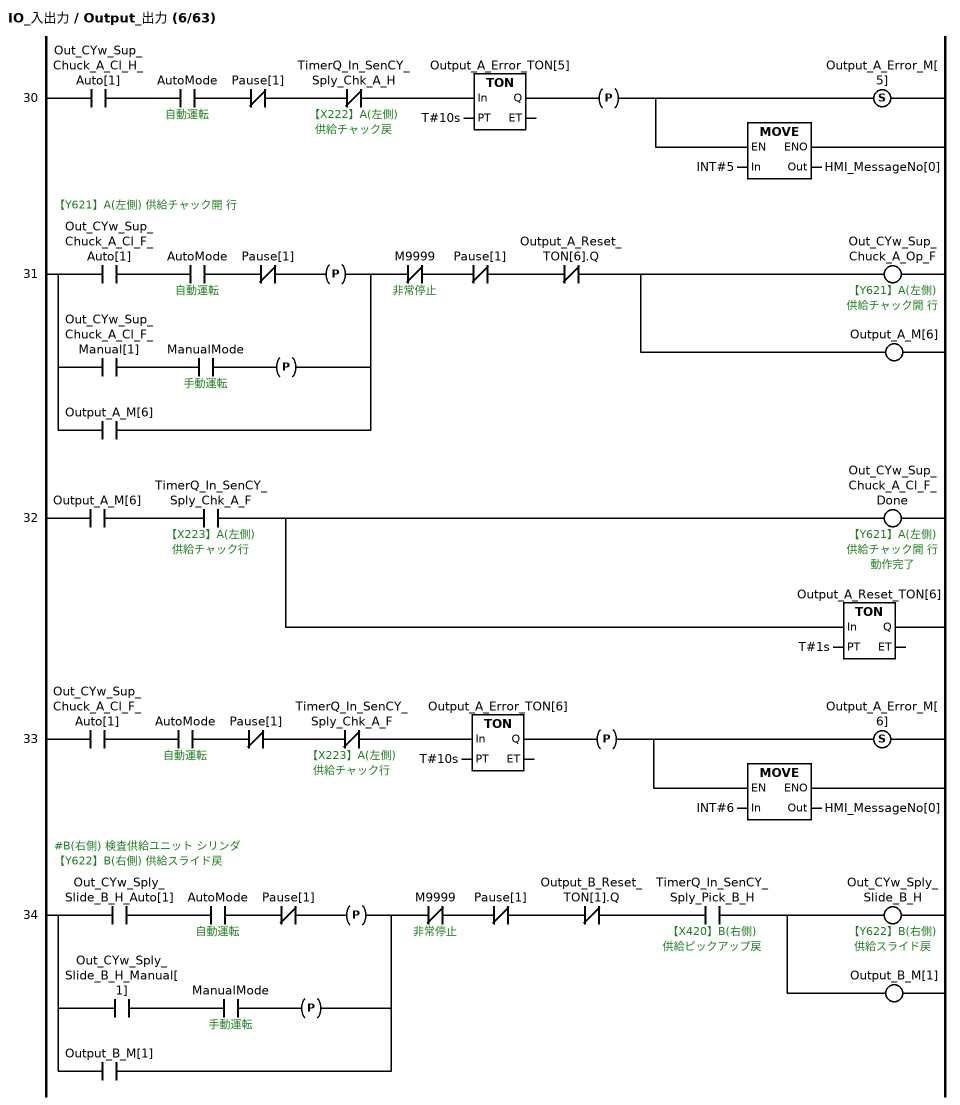
(* [picture p74: IO_入出力 / Output_出力, rungs 30-34] *)
(* Rung 30 *)
Output_A_Error_TON[5](In := Out_CYw_Sup_Chuck_A_Cl_H_Auto[1] AND AutoMode AND NOT Pause[1] AND NOT TimerQ_In_SenCY_Sply_Chk_A_H, PT := T#10s);
_e20(CLK := Output_A_Error_TON[5].Q);
IF _e20.Q THEN
    Output_A_Error_M[5] := TRUE;
    HMI_MessageNo[0] := INT#5;
END_IF;
(* Rung 31: 【Y621】A(左側) 供給チャック開 行 *)
_e21(CLK := Out_CYw_Sup_Chuck_A_Cl_F_Auto[1] AND AutoMode AND NOT Pause[1]);
_e22(CLK := Out_CYw_Sup_Chuck_A_Cl_F_Manual[1] AND ManualMode);
_p23 := (_e21.Q OR _e22.Q OR Output_A_M[6]) AND NOT M9999 AND NOT Pause[1] AND NOT Output_A_Reset_TON[6].Q;
Out_CYw_Sup_Chuck_A_Op_F := _p23;
Output_A_M[6] := _p23;
(* Rung 32 *)
Out_CYw_Sup_Chuck_A_Cl_F_Done := Output_A_M[6] AND TimerQ_In_SenCY_Sply_Chk_A_F;
Output_A_Reset_TON[6](In := Output_A_M[6] AND TimerQ_In_SenCY_Sply_Chk_A_F, PT := T#1s);
(* Rung 33 *)
Output_A_Error_TON[6](In := Out_CYw_Sup_Chuck_A_Cl_F_Auto[1] AND AutoMode AND NOT Pause[1] AND NOT TimerQ_In_SenCY_Sply_Chk_A_F, PT := T#10s);
_e24(CLK := Output_A_Error_TON[6].Q);
IF _e24.Q THEN
    Output_A_Error_M[6] := TRUE;
    HMI_MessageNo[0] := INT#6;
END_IF;
(* Rung 34: #B(右側) 検査供給ユニット シリンダ / 【Y622】B(右側) 供給スライド戻 *)
_e25(CLK := Out_CYw_Sply_Slide_B_H_Auto[1] AND AutoMode AND NOT Pause[1]);
_e26(CLK := Out_CYw_Sply_Slide_B_H_Manual[1] AND ManualMode);
_p27 := (_e25.Q OR _e26.Q OR Output_B_M[1]) AND NOT M9999 AND NOT Pause[1] AND NOT Output_B_Reset_TON[1].Q AND TimerQ_In_SenCY_Sply_Pick_B_H;
Out_CYw_Sply_Slide_B_H := _p27;
Output_B_M[1] := _p27;

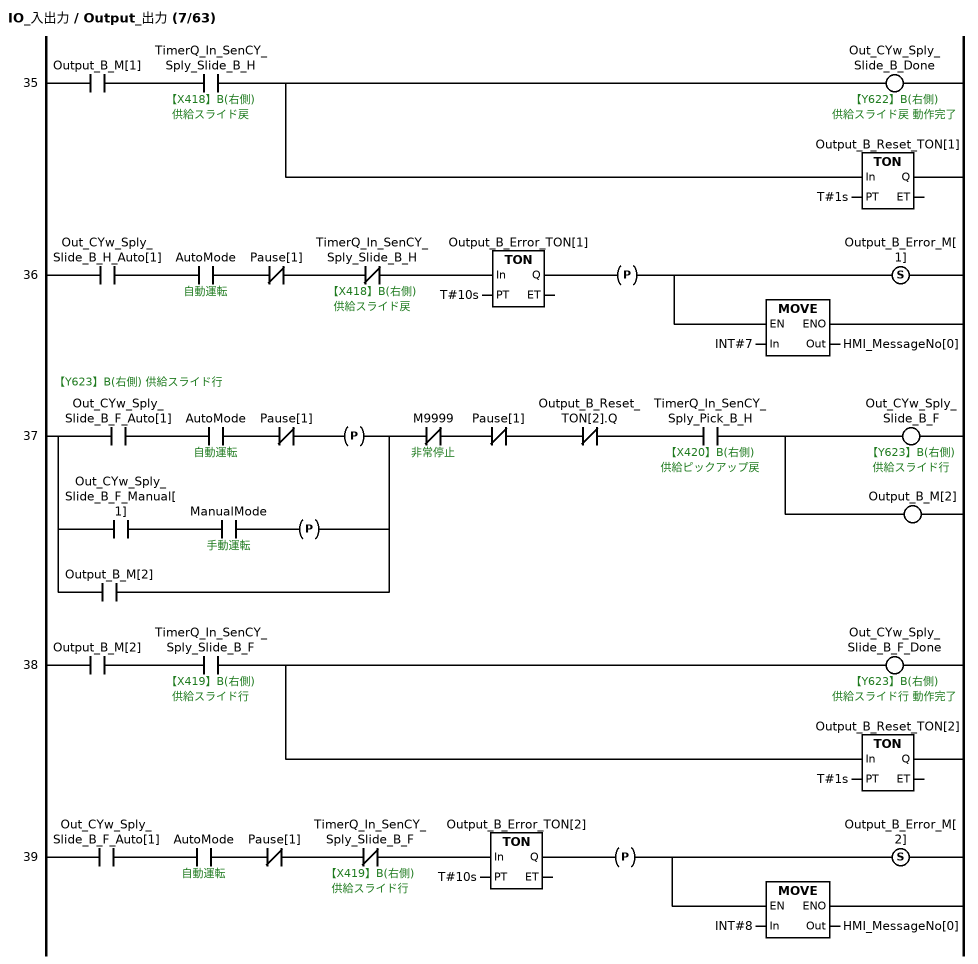
(* Rung 35 *)
Out_CYw_Sply_Slide_B_Done := Output_B_M[1] AND TimerQ_In_SenCY_Sply_Slide_B_H;
Output_B_Reset_TON[1](In := Output_B_M[1] AND TimerQ_In_SenCY_Sply_Slide_B_H, PT := T#1s);
(* Rung 36 *)
Output_B_Error_TON[1](In := Out_CYw_Sply_Slide_B_H_Auto[1] AND AutoMode AND NOT Pause[1] AND NOT TimerQ_In_SenCY_Sply_Slide_B_H, PT := T#10s);
_e28(CLK := Output_B_Error_TON[1].Q);
IF _e28.Q THEN
    Output_B_Error_M[1] := TRUE;
    HMI_MessageNo[0] := INT#7;
END_IF;
(* Rung 37: 【Y623】B(右側) 供給スライド行 *)
_e29(CLK := Out_CYw_Sply_Slide_B_F_Auto[1] AND AutoMode AND NOT Pause[1]);
_e30(CLK := Out_CYw_Sply_Slide_B_F_Manual[1] AND ManualMode);
_p31 := (_e29.Q OR _e30.Q OR Output_B_M[2]) AND NOT M9999 AND NOT Pause[1] AND NOT Output_B_Reset_TON[2].Q AND TimerQ_In_SenCY_Sply_Pick_B_H;
Out_CYw_Sply_Slide_B_F := _p31;
Output_B_M[2] := _p31;
(* Rung 38 *)
Out_CYw_Sply_Slide_B_F_Done := Output_B_M[2] AND TimerQ_In_SenCY_Sply_Slide_B_F;
Output_B_Reset_TON[2](In := Output_B_M[2] AND TimerQ_In_SenCY_Sply_Slide_B_F, PT := T#1s);
(* Rung 39 *)
Output_B_Error_TON[2](In := Out_CYw_Sply_Slide_B_F_Auto[1] AND AutoMode AND NOT Pause[1] AND NOT TimerQ_In_SenCY_Sply_Slide_B_F, PT := T#10s);
_e32(CLK := Output_B_Error_TON[2].Q);
IF _e32.Q THEN
    Output_B_Error_M[2] := TRUE;
    HMI_MessageNo[0] := INT#8;
END_IF;

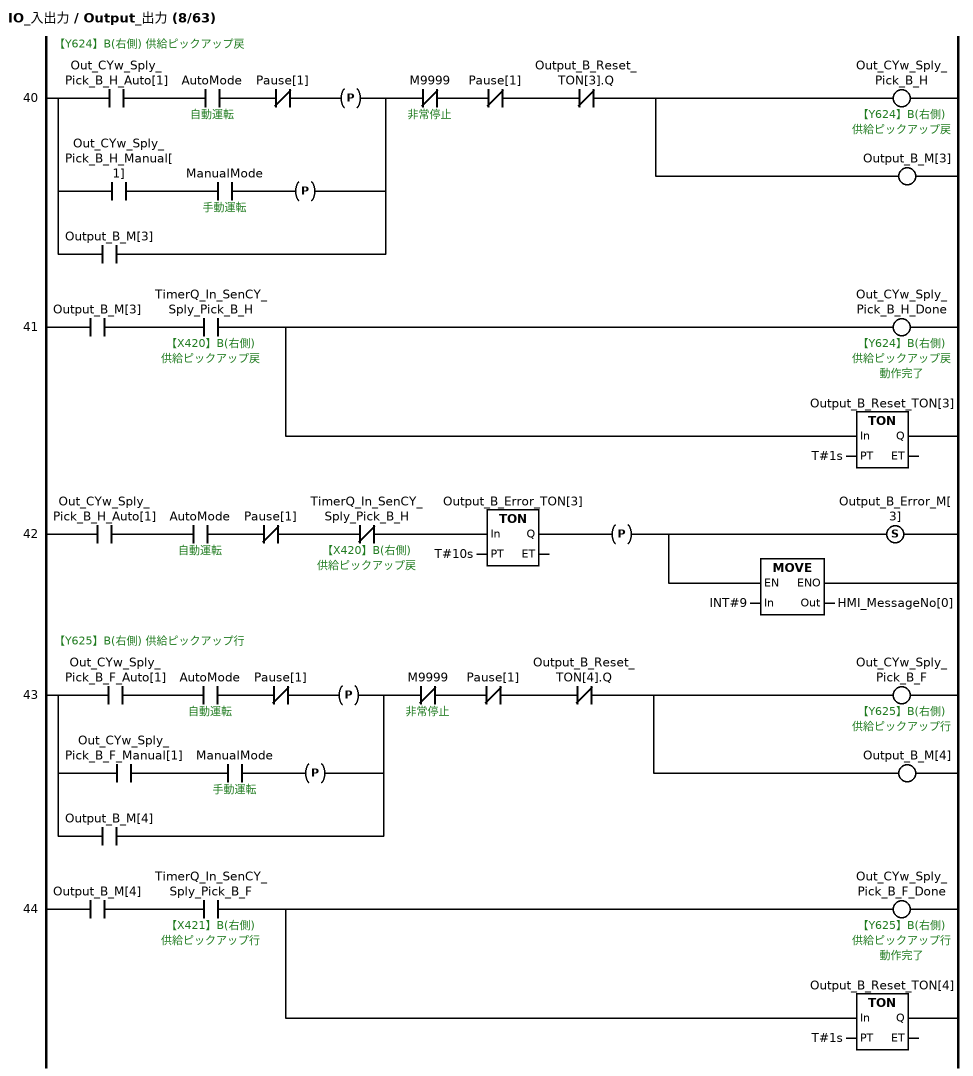
(* Rung 40: 【Y624】B(右側) 供給ピックアップ戻 *)
_e33(CLK := Out_CYw_Sply_Pick_B_H_Auto[1] AND AutoMode AND NOT Pause[1]);
_e34(CLK := Out_CYw_Sply_Pick_B_H_Manual[1] AND ManualMode);
_p35 := (_e33.Q OR _e34.Q OR Output_B_M[3]) AND NOT M9999 AND NOT Pause[1] AND NOT Output_B_Reset_TON[3].Q;
Out_CYw_Sply_Pick_B_H := _p35;
Output_B_M[3] := _p35;
(* Rung 41 *)
Out_CYw_Sply_Pick_B_H_Done := Output_B_M[3] AND TimerQ_In_SenCY_Sply_Pick_B_H;
Output_B_Reset_TON[3](In := Output_B_M[3] AND TimerQ_In_SenCY_Sply_Pick_B_H, PT := T#1s);
(* Rung 42 *)
Output_B_Error_TON[3](In := Out_CYw_Sply_Pick_B_H_Auto[1] AND AutoMode AND NOT Pause[1] AND NOT TimerQ_In_SenCY_Sply_Pick_B_H, PT := T#10s);
_e36(CLK := Output_B_Error_TON[3].Q);
IF _e36.Q THEN
    Output_B_Error_M[3] := TRUE;
    HMI_MessageNo[0] := INT#9;
END_IF;
(* Rung 43: 【Y625】B(右側) 供給ピックアップ行 *)
_e37(CLK := Out_CYw_Sply_Pick_B_F_Auto[1] AND AutoMode AND NOT Pause[1]);
_e38(CLK := Out_CYw_Sply_Pick_B_F_Manual[1] AND ManualMode);
_p39 := (_e37.Q OR _e38.Q OR Output_B_M[4]) AND NOT M9999 AND NOT Pause[1] AND NOT Output_B_Reset_TON[4].Q;
Out_CYw_Sply_Pick_B_F := _p39;
Output_B_M[4] := _p39;
(* Rung 44 *)
Out_CYw_Sply_Pick_B_F_Done := Output_B_M[4] AND TimerQ_In_SenCY_Sply_Pick_B_F;
Output_B_Reset_TON[4](In := Output_B_M[4] AND TimerQ_In_SenCY_Sply_Pick_B_F, PT := T#1s);

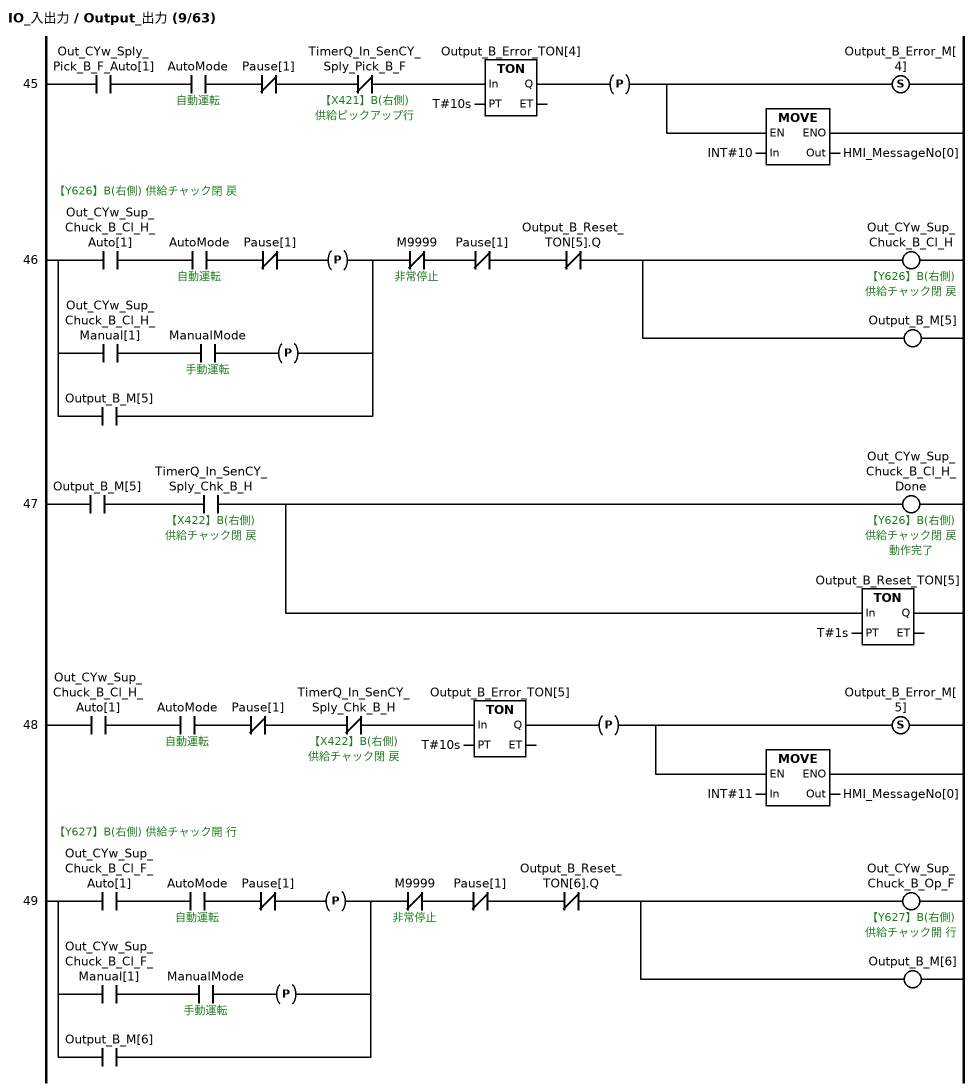
(* Rung 45 *)
Output_B_Error_TON[4](In := Out_CYw_Sply_Pick_B_F_Auto[1] AND AutoMode AND NOT Pause[1] AND NOT TimerQ_In_SenCY_Sply_Pick_B_F, PT := T#10s);
_e40(CLK := Output_B_Error_TON[4].Q);
IF _e40.Q THEN
    Output_B_Error_M[4] := TRUE;
    HMI_MessageNo[0] := INT#10;
END_IF;
(* Rung 46: 【Y626】B(右側) 供給チャック閉 戻 *)
_e41(CLK := Out_CYw_Sup_Chuck_B_Cl_H_Auto[1] AND AutoMode AND NOT Pause[1]);
_e42(CLK := Out_CYw_Sup_Chuck_B_Cl_H_Manual[1] AND ManualMode);
_p43 := (_e41.Q OR _e42.Q OR Output_B_M[5]) AND NOT M9999 AND NOT Pause[1] AND NOT Output_B_Reset_TON[5].Q;
Out_CYw_Sup_Chuck_B_Cl_H := _p43;
Output_B_M[5] := _p43;
(* Rung 47 *)
Out_CYw_Sup_Chuck_B_Cl_H_Done := Output_B_M[5] AND TimerQ_In_SenCY_Sply_Chk_B_H;
Output_B_Reset_TON[5](In := Output_B_M[5] AND TimerQ_In_SenCY_Sply_Chk_B_H, PT := T#1s);
(* Rung 48 *)
Output_B_Error_TON[5](In := Out_CYw_Sup_Chuck_B_Cl_H_Auto[1] AND AutoMode AND NOT Pause[1] AND NOT TimerQ_In_SenCY_Sply_Chk_B_H, PT := T#10s);
_e44(CLK := Output_B_Error_TON[5].Q);
IF _e44.Q THEN
    Output_B_Error_M[5] := TRUE;
    HMI_MessageNo[0] := INT#11;
END_IF;
(* Rung 49: 【Y627】B(右側) 供給チャック開 行 *)
_e45(CLK := Out_CYw_Sup_Chuck_B_Cl_F_Auto[1] AND AutoMode AND NOT Pause[1]);
_e46(CLK := Out_CYw_Sup_Chuck_B_Cl_F_Manual[1] AND ManualMode);
_p47 := (_e45.Q OR _e46.Q OR Output_B_M[6]) AND NOT M9999 AND NOT Pause[1] AND NOT Output_B_Reset_TON[6].Q;
Out_CYw_Sup_Chuck_B_Op_F := _p47;
Output_B_M[6] := _p47;

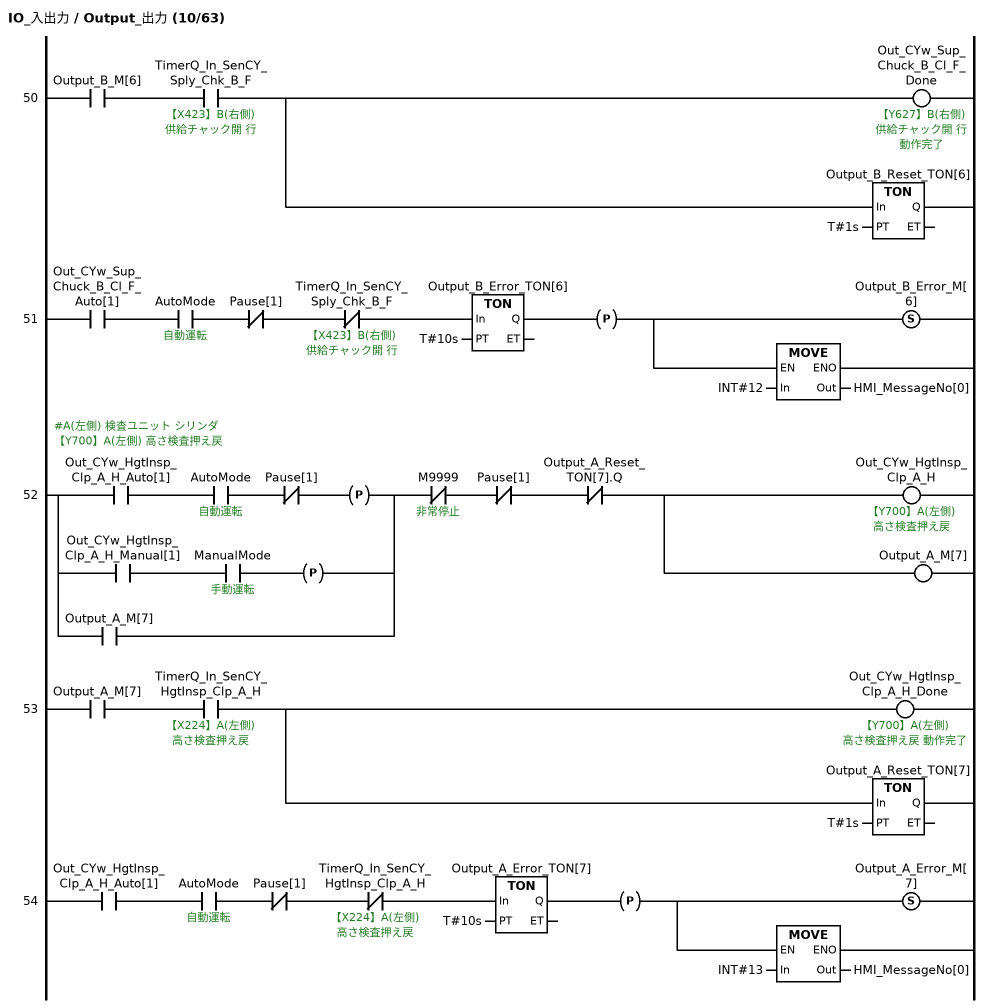
(* Rung 50 *)
Out_CYw_Sup_Chuck_B_Cl_F_Done := Output_B_M[6] AND TimerQ_In_SenCY_Sply_Chk_B_F;
Output_B_Reset_TON[6](In := Output_B_M[6] AND TimerQ_In_SenCY_Sply_Chk_B_F, PT := T#1s);
(* Rung 51 *)
Output_B_Error_TON[6](In := Out_CYw_Sup_Chuck_B_Cl_F_Auto[1] AND AutoMode AND NOT Pause[1] AND NOT TimerQ_In_SenCY_Sply_Chk_B_F, PT := T#10s);
_e48(CLK := Output_B_Error_TON[6].Q);
IF _e48.Q THEN
    Output_B_Error_M[6] := TRUE;
    HMI_MessageNo[0] := INT#12;
END_IF;
(* Rung 52: #A(左側) 検査ユニット シリンダ / 【Y700】A(左側) 高さ検査押え戻 *)
_e49(CLK := Out_CYw_HgtInsp_Clp_A_H_Auto[1] AND AutoMode AND NOT Pause[1]);
_e50(CLK := Out_CYw_HgtInsp_Clp_A_H_Manual[1] AND ManualMode);
_p51 := (_e49.Q OR _e50.Q OR Output_A_M[7]) AND NOT M9999 AND NOT Pause[1] AND NOT Output_A_Reset_TON[7].Q;
Out_CYw_HgtInsp_Clp_A_H := _p51;
Output_A_M[7] := _p51;
(* Rung 53 *)
_p52 := Output_A_M[7] AND TimerQ_In_SenCY_HgtInsp_Clp_A_H;
Out_CYw_HgtInsp_Clp_A_H_Done := _p52;
Output_A_Reset_TON[7](In := _p52, PT := T#1s);
(* Rung 54 *)
Output_A_Error_TON[7](In := Out_CYw_HgtInsp_Clp_A_H_Auto[1] AND AutoMode AND NOT Pause[1] AND NOT TimerQ_In_SenCY_HgtInsp_Clp_A_H, PT := T#10s);
_e53(CLK := Output_A_Error_TON[7].Q);
IF _e53.Q THEN
    Output_A_Error_M[7] := TRUE;
    HMI_MessageNo[0] := INT#13;
END_IF;

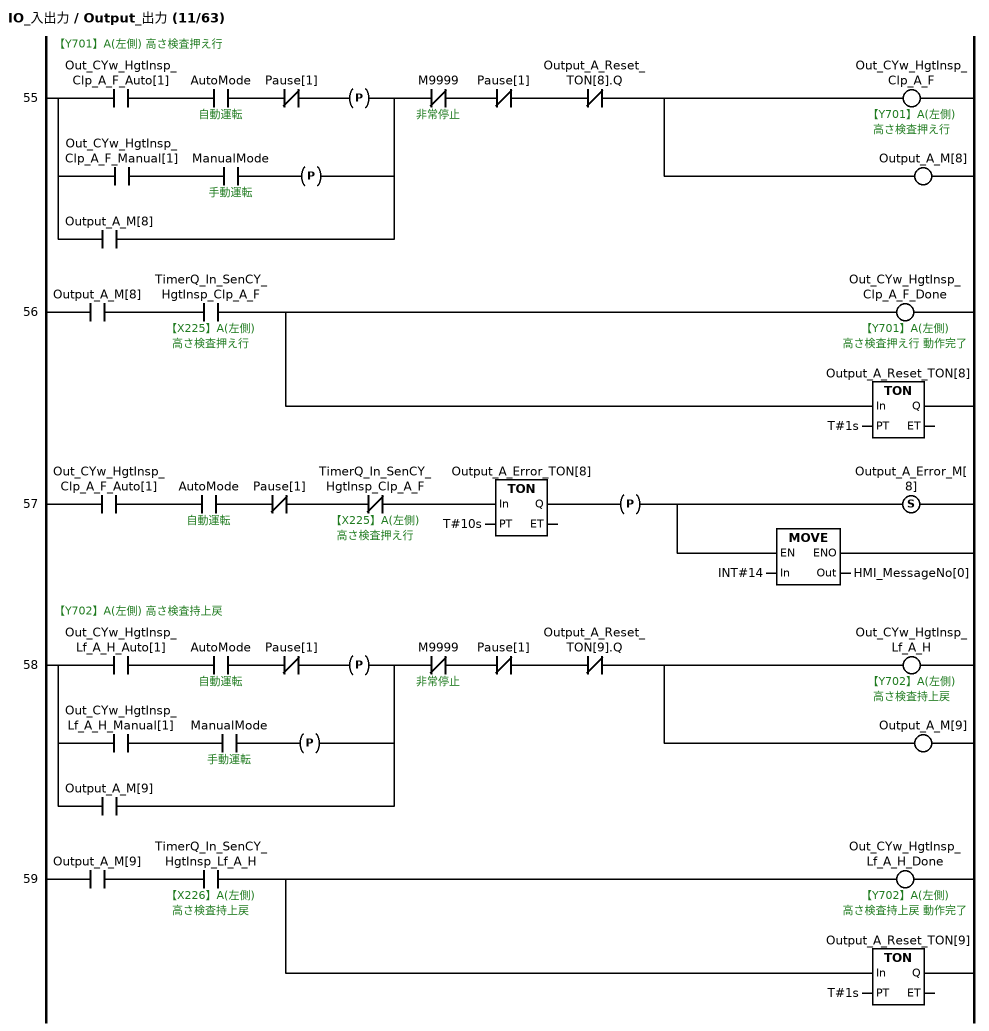
(* Rung 55: 【Y701】A(左側) 高さ検査押え行 *)
_e54(CLK := Out_CYw_HgtInsp_Clp_A_F_Auto[1] AND AutoMode AND NOT Pause[1]);
_e55(CLK := Out_CYw_HgtInsp_Clp_A_F_Manual[1] AND ManualMode);
_p56 := (_e54.Q OR _e55.Q OR Output_A_M[8]) AND NOT M9999 AND NOT Pause[1] AND NOT Output_A_Reset_TON[8].Q;
Out_CYw_HgtInsp_Clp_A_F := _p56;
Output_A_M[8] := _p56;
(* Rung 56 *)
_p57 := Output_A_M[8] AND TimerQ_In_SenCY_HgtInsp_Clp_A_F;
Out_CYw_HgtInsp_Clp_A_F_Done := _p57;
Output_A_Reset_TON[8](In := _p57, PT := T#1s);
(* Rung 57 *)
Output_A_Error_TON[8](In := Out_CYw_HgtInsp_Clp_A_F_Auto[1] AND AutoMode AND NOT Pause[1] AND NOT TimerQ_In_SenCY_HgtInsp_Clp_A_F, PT := T#10s);
_e58(CLK := Output_A_Error_TON[8].Q);
IF _e58.Q THEN
    Output_A_Error_M[8] := TRUE;
    HMI_MessageNo[0] := INT#14;
END_IF;
(* Rung 58: 【Y702】A(左側) 高さ検査持上戻 *)
_e59(CLK := Out_CYw_HgtInsp_Lf_A_H_Auto[1] AND AutoMode AND NOT Pause[1]);
_e60(CLK := Out_CYw_HgtInsp_Lf_A_H_Manual[1] AND ManualMode);
_p61 := (_e59.Q OR _e60.Q OR Output_A_M[9]) AND NOT M9999 AND NOT Pause[1] AND NOT Output_A_Reset_TON[9].Q;
Out_CYw_HgtInsp_Lf_A_H := _p61;
Output_A_M[9] := _p61;
(* Rung 59 *)
Out_CYw_HgtInsp_Lf_A_H_Done := Output_A_M[9] AND TimerQ_In_SenCY_HgtInsp_Lf_A_H;
Output_A_Reset_TON[9](In := Output_A_M[9] AND TimerQ_In_SenCY_HgtInsp_Lf_A_H, PT := T#1s);

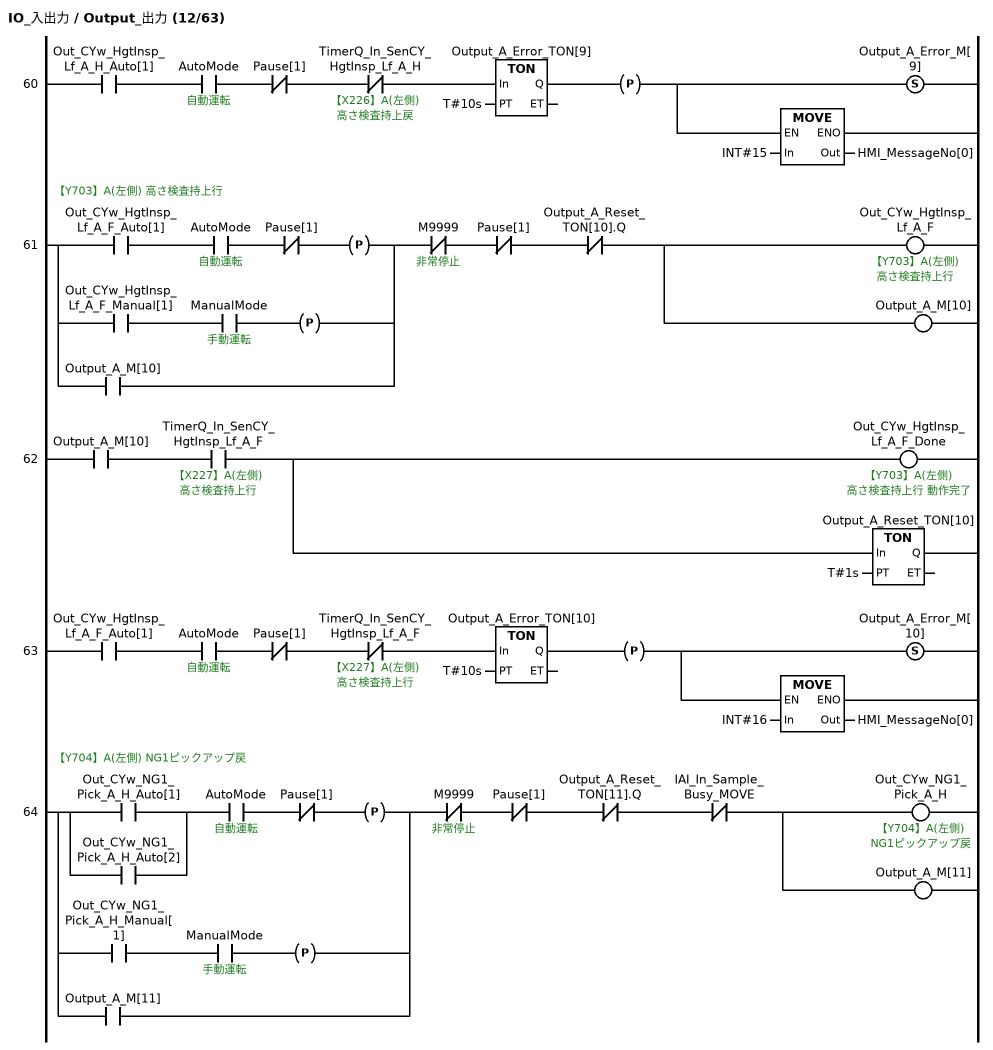
(* Rung 60 *)
Output_A_Error_TON[9](In := Out_CYw_HgtInsp_Lf_A_H_Auto[1] AND AutoMode AND NOT Pause[1] AND NOT TimerQ_In_SenCY_HgtInsp_Lf_A_H, PT := T#10s);
_e62(CLK := Output_A_Error_TON[9].Q);
IF _e62.Q THEN
    Output_A_Error_M[9] := TRUE;
    HMI_MessageNo[0] := INT#15;
END_IF;
(* Rung 61: 【Y703】A(左側) 高さ検査持上行 *)
_e63(CLK := Out_CYw_HgtInsp_Lf_A_F_Auto[1] AND AutoMode AND NOT Pause[1]);
_e64(CLK := Out_CYw_HgtInsp_Lf_A_F_Manual[1] AND ManualMode);
_p65 := (_e63.Q OR _e64.Q OR Output_A_M[10]) AND NOT M9999 AND NOT Pause[1] AND NOT Output_A_Reset_TON[10].Q;
Out_CYw_HgtInsp_Lf_A_F := _p65;
Output_A_M[10] := _p65;
(* Rung 62 *)
_p66 := Output_A_M[10] AND TimerQ_In_SenCY_HgtInsp_Lf_A_F;
Out_CYw_HgtInsp_Lf_A_F_Done := _p66;
Output_A_Reset_TON[10](In := _p66, PT := T#1s);
(* Rung 63 *)
Output_A_Error_TON[10](In := Out_CYw_HgtInsp_Lf_A_F_Auto[1] AND AutoMode AND NOT Pause[1] AND NOT TimerQ_In_SenCY_HgtInsp_Lf_A_F, PT := T#10s);
_e67(CLK := Output_A_Error_TON[10].Q);
IF _e67.Q THEN
    Output_A_Error_M[10] := TRUE;
    HMI_MessageNo[0] := INT#16;
END_IF;
(* Rung 64: 【Y704】A(左側) NG1ピックアップ戻 *)
_e68(CLK := (Out_CYw_NG1_Pick_A_H_Auto[1] OR Out_CYw_NG1_Pick_A_H_Auto[2]) AND AutoMode AND NOT Pause[1]);
_e69(CLK := Out_CYw_NG1_Pick_A_H_Manual[1] AND ManualMode);
_p70 := (_e68.Q OR _e69.Q OR Output_A_M[11]) AND NOT M9999 AND NOT Pause[1] AND NOT Output_A_Reset_TON[11].Q AND NOT IAI_In_Sample_Busy_MOVE;
Out_CYw_NG1_Pick_A_H := _p70;
Output_A_M[11] := _p70;

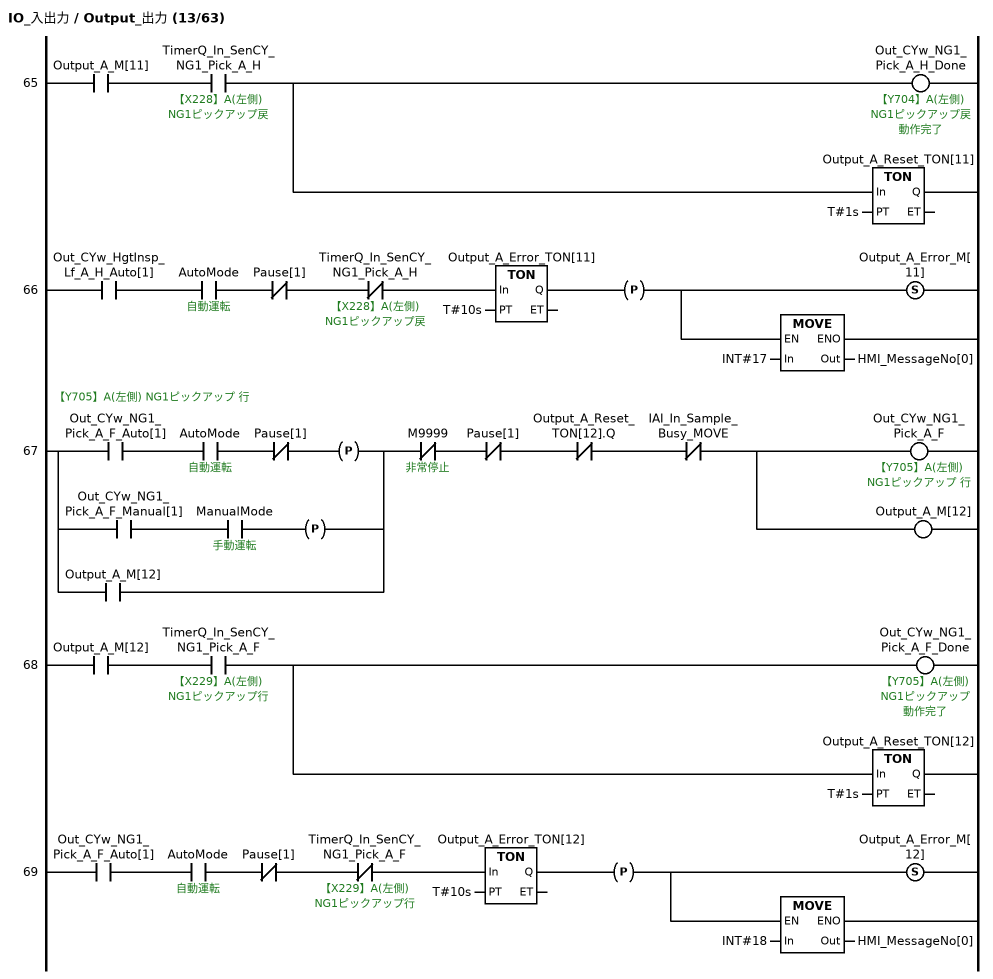
(* Rung 65 *)
Out_CYw_NG1_Pick_A_H_Done := Output_A_M[11] AND TimerQ_In_SenCY_NG1_Pick_A_H;
Output_A_Reset_TON[11](In := Output_A_M[11] AND TimerQ_In_SenCY_NG1_Pick_A_H, PT := T#1s);
(* Rung 66 *)
Output_A_Error_TON[11](In := Out_CYw_HgtInsp_Lf_A_H_Auto[1] AND AutoMode AND NOT Pause[1] AND NOT TimerQ_In_SenCY_NG1_Pick_A_H, PT := T#10s);
_e71(CLK := Output_A_Error_TON[11].Q);
IF _e71.Q THEN
    Output_A_Error_M[11] := TRUE;
    HMI_MessageNo[0] := INT#17;
END_IF;
(* Rung 67: 【Y705】A(左側) NG1ピックアップ 行 *)
_e72(CLK := Out_CYw_NG1_Pick_A_F_Auto[1] AND AutoMode AND NOT Pause[1]);
_e73(CLK := Out_CYw_NG1_Pick_A_F_Manual[1] AND ManualMode);
_p74 := (_e72.Q OR _e73.Q OR Output_A_M[12]) AND NOT M9999 AND NOT Pause[1] AND NOT Output_A_Reset_TON[12].Q AND NOT IAI_In_Sample_Busy_MOVE;
Out_CYw_NG1_Pick_A_F := _p74;
Output_A_M[12] := _p74;
(* Rung 68 *)
Out_CYw_NG1_Pick_A_F_Done := Output_A_M[12] AND TimerQ_In_SenCY_NG1_Pick_A_F;
Output_A_Reset_TON[12](In := Output_A_M[12] AND TimerQ_In_SenCY_NG1_Pick_A_F, PT := T#1s);
(* Rung 69 *)
Output_A_Error_TON[12](In := Out_CYw_NG1_Pick_A_F_Auto[1] AND AutoMode AND NOT Pause[1] AND NOT TimerQ_In_SenCY_NG1_Pick_A_F, PT := T#10s);
_e75(CLK := Output_A_Error_TON[12].Q);
IF _e75.Q THEN
    Output_A_Error_M[12] := TRUE;
    HMI_MessageNo[0] := INT#18;
END_IF;

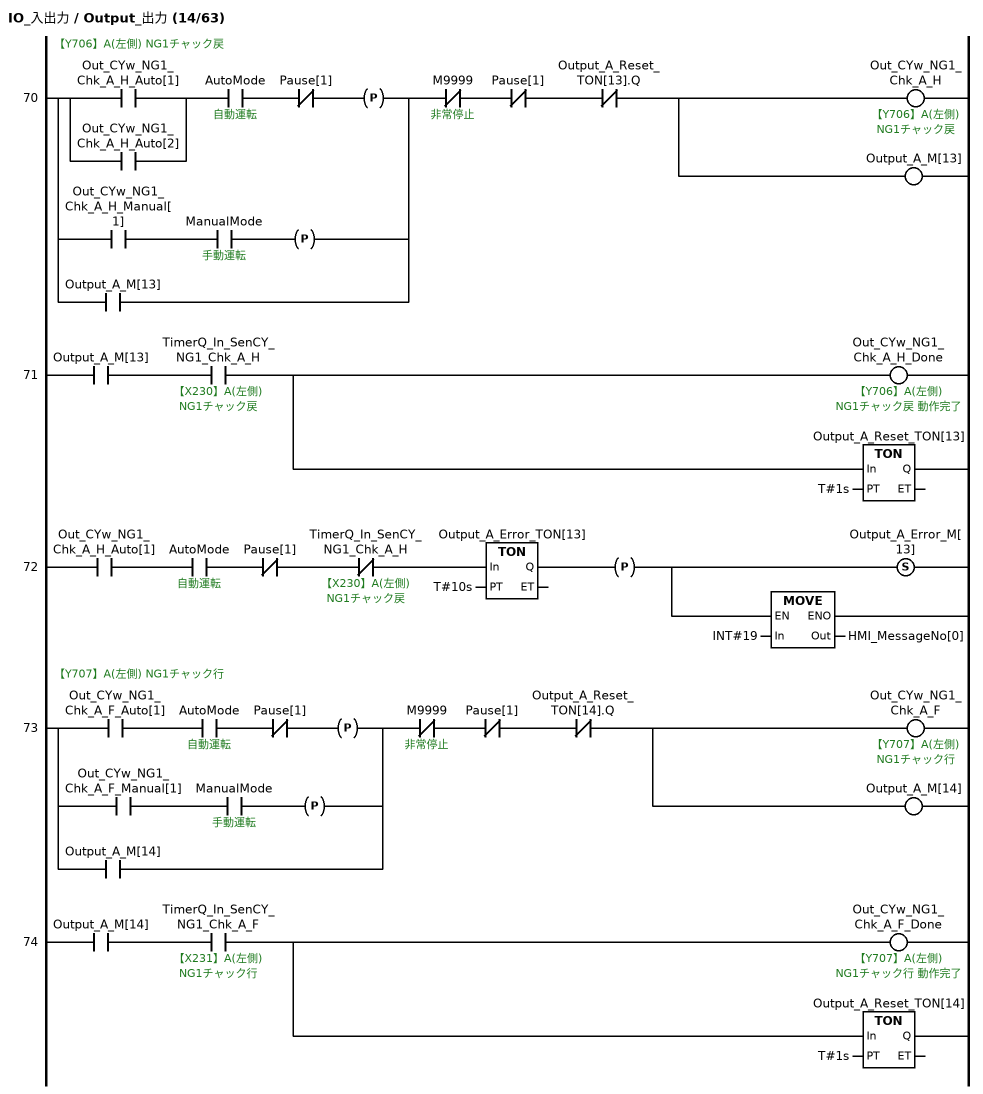
(* Rung 70: 【Y706】A(左側) NG1チャック戻 *)
_e76(CLK := (Out_CYw_NG1_Chk_A_H_Auto[1] OR Out_CYw_NG1_Chk_A_H_Auto[2]) AND AutoMode AND NOT Pause[1]);
_e77(CLK := Out_CYw_NG1_Chk_A_H_Manual[1] AND ManualMode);
_p78 := (_e76.Q OR _e77.Q OR Output_A_M[13]) AND NOT M9999 AND NOT Pause[1] AND NOT Output_A_Reset_TON[13].Q;
Out_CYw_NG1_Chk_A_H := _p78;
Output_A_M[13] := _p78;
(* Rung 71 *)
Out_CYw_NG1_Chk_A_H_Done := Output_A_M[13] AND TimerQ_In_SenCY_NG1_Chk_A_H;
Output_A_Reset_TON[13](In := Output_A_M[13] AND TimerQ_In_SenCY_NG1_Chk_A_H, PT := T#1s);
(* Rung 72 *)
Output_A_Error_TON[13](In := Out_CYw_NG1_Chk_A_H_Auto[1] AND AutoMode AND NOT Pause[1] AND NOT TimerQ_In_SenCY_NG1_Chk_A_H, PT := T#10s);
_e79(CLK := Output_A_Error_TON[13].Q);
IF _e79.Q THEN
    Output_A_Error_M[13] := TRUE;
    HMI_MessageNo[0] := INT#19;
END_IF;
(* Rung 73: 【Y707】A(左側) NG1チャック行 *)
_e80(CLK := Out_CYw_NG1_Chk_A_F_Auto[1] AND AutoMode AND NOT Pause[1]);
_e81(CLK := Out_CYw_NG1_Chk_A_F_Manual[1] AND ManualMode);
_p82 := (_e80.Q OR _e81.Q OR Output_A_M[14]) AND NOT M9999 AND NOT Pause[1] AND NOT Output_A_Reset_TON[14].Q;
Out_CYw_NG1_Chk_A_F := _p82;
Output_A_M[14] := _p82;
(* Rung 74 *)
Out_CYw_NG1_Chk_A_F_Done := Output_A_M[14] AND TimerQ_In_SenCY_NG1_Chk_A_F;
Output_A_Reset_TON[14](In := Output_A_M[14] AND TimerQ_In_SenCY_NG1_Chk_A_F, PT := T#1s);

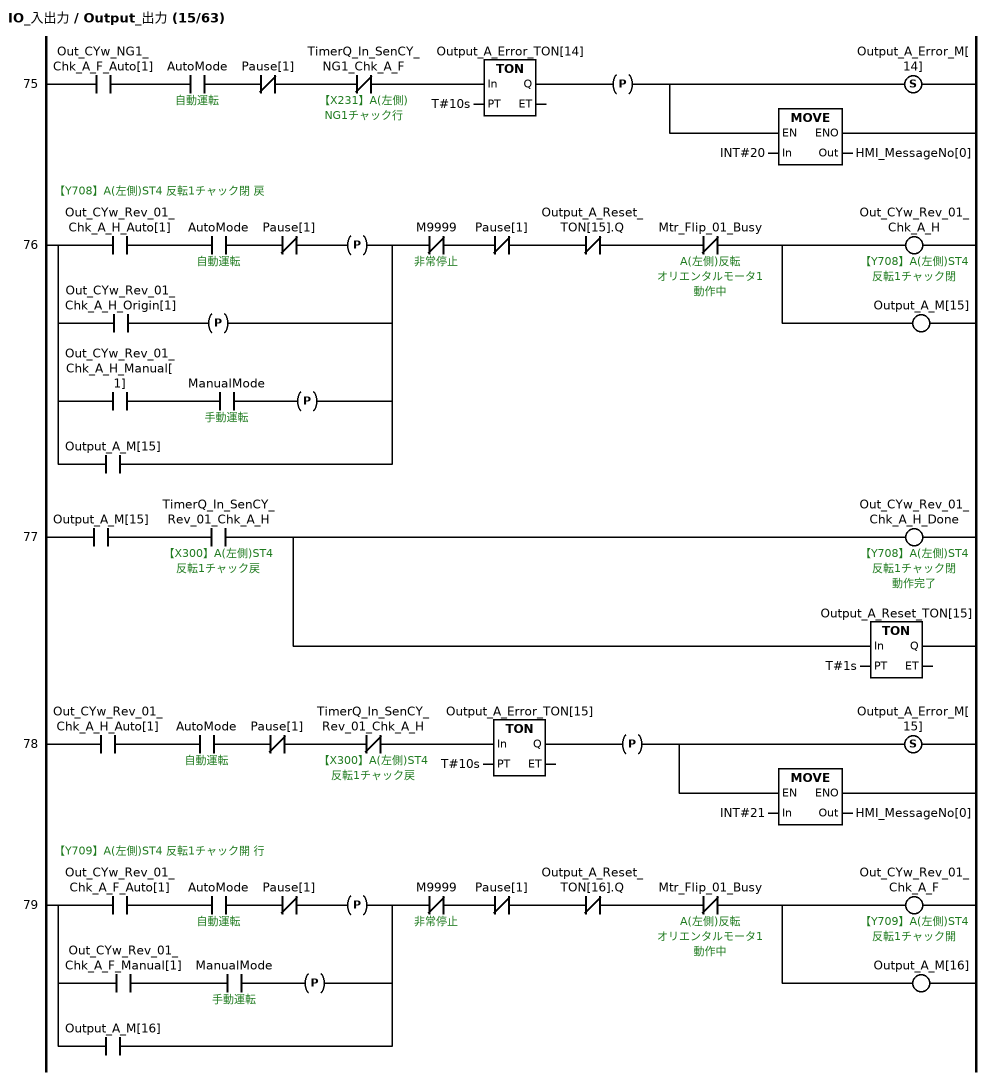
(* Rung 75 *)
Output_A_Error_TON[14](In := Out_CYw_NG1_Chk_A_F_Auto[1] AND AutoMode AND NOT Pause[1] AND NOT TimerQ_In_SenCY_NG1_Chk_A_F, PT := T#10s);
_e83(CLK := Output_A_Error_TON[14].Q);
IF _e83.Q THEN
    Output_A_Error_M[14] := TRUE;
    HMI_MessageNo[0] := INT#20;
END_IF;
(* Rung 76: 【Y708】A(左側)ST4 反転1チャック閉 戻 *)
_e84(CLK := Out_CYw_Rev_01_Chk_A_H_Auto[1] AND AutoMode AND NOT Pause[1]);
_e85(CLK := Out_CYw_Rev_01_Chk_A_H_Origin[1]);
_e86(CLK := Out_CYw_Rev_01_Chk_A_H_Manual[1] AND ManualMode);
_p87 := (_e84.Q OR _e85.Q OR _e86.Q OR Output_A_M[15]) AND NOT M9999 AND NOT Pause[1] AND NOT Output_A_Reset_TON[15].Q AND NOT Mtr_Flip_01_Busy;
Out_CYw_Rev_01_Chk_A_H := _p87;
Output_A_M[15] := _p87;
(* Rung 77 *)
_p88 := Output_A_M[15] AND TimerQ_In_SenCY_Rev_01_Chk_A_H;
Out_CYw_Rev_01_Chk_A_H_Done := _p88;
Output_A_Reset_TON[15](In := _p88, PT := T#1s);
(* Rung 78 *)
Output_A_Error_TON[15](In := Out_CYw_Rev_01_Chk_A_H_Auto[1] AND AutoMode AND NOT Pause[1] AND NOT TimerQ_In_SenCY_Rev_01_Chk_A_H, PT := T#10s);
_e89(CLK := Output_A_Error_TON[15].Q);
IF _e89.Q THEN
    Output_A_Error_M[15] := TRUE;
    HMI_MessageNo[0] := INT#21;
END_IF;
(* Rung 79: 【Y709】A(左側)ST4 反転1チャック開 行 *)
_e90(CLK := Out_CYw_Rev_01_Chk_A_F_Auto[1] AND AutoMode AND NOT Pause[1]);
_e91(CLK := Out_CYw_Rev_01_Chk_A_F_Manual[1] AND ManualMode);
_p92 := (_e90.Q OR _e91.Q OR Output_A_M[16]) AND NOT M9999 AND NOT Pause[1] AND NOT Output_A_Reset_TON[16].Q AND NOT Mtr_Flip_01_Busy;
Out_CYw_Rev_01_Chk_A_F := _p92;
Output_A_M[16] := _p92;

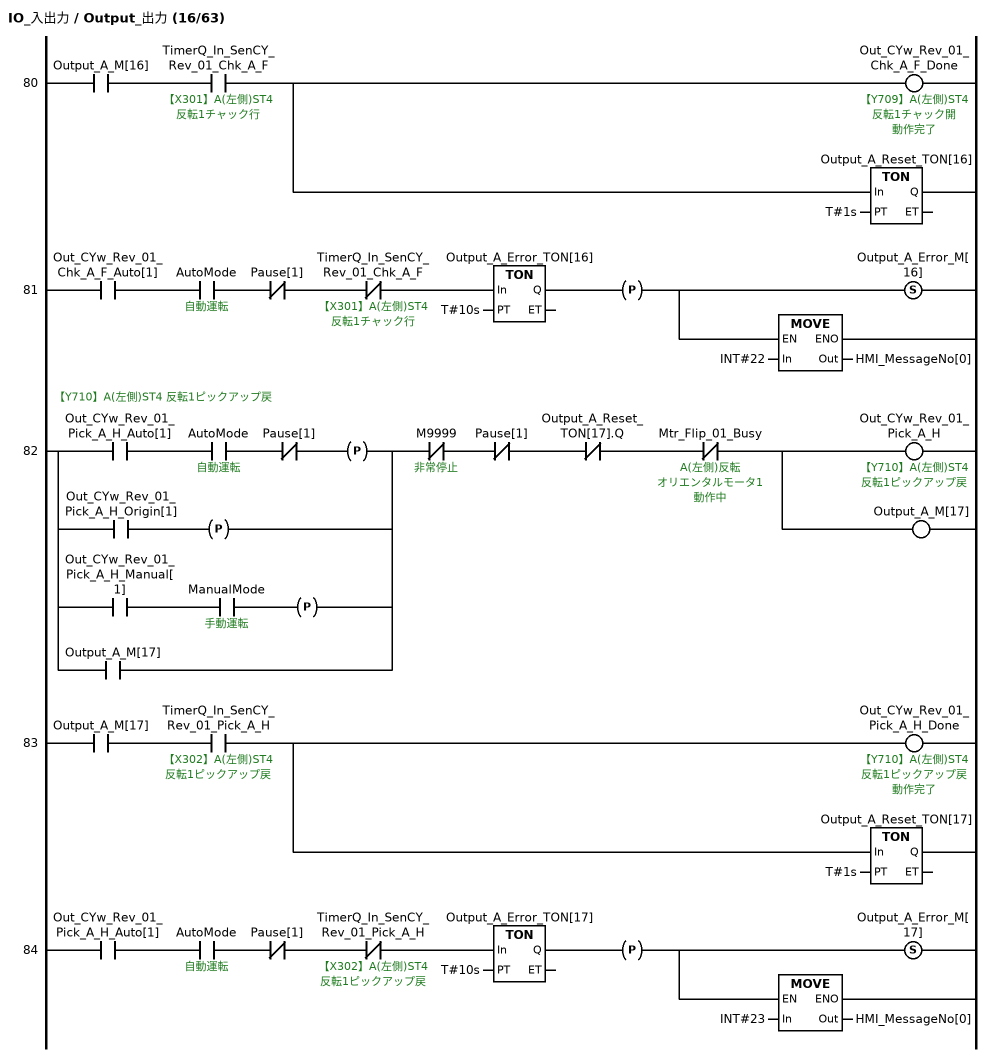
(* Rung 80 *)
_p93 := Output_A_M[16] AND TimerQ_In_SenCY_Rev_01_Chk_A_F;
Out_CYw_Rev_01_Chk_A_F_Done := _p93;
Output_A_Reset_TON[16](In := _p93, PT := T#1s);
(* Rung 81 *)
Output_A_Error_TON[16](In := Out_CYw_Rev_01_Chk_A_F_Auto[1] AND AutoMode AND NOT Pause[1] AND NOT TimerQ_In_SenCY_Rev_01_Chk_A_F, PT := T#10s);
_e94(CLK := Output_A_Error_TON[16].Q);
IF _e94.Q THEN
    Output_A_Error_M[16] := TRUE;
    HMI_MessageNo[0] := INT#22;
END_IF;
(* Rung 82: 【Y710】A(左側)ST4 反転1ピックアップ戻 *)
_e95(CLK := Out_CYw_Rev_01_Pick_A_H_Auto[1] AND AutoMode AND NOT Pause[1]);
_e96(CLK := Out_CYw_Rev_01_Pick_A_H_Origin[1]);
_e97(CLK := Out_CYw_Rev_01_Pick_A_H_Manual[1] AND ManualMode);
_p98 := (_e95.Q OR _e96.Q OR _e97.Q OR Output_A_M[17]) AND NOT M9999 AND NOT Pause[1] AND NOT Output_A_Reset_TON[17].Q AND NOT Mtr_Flip_01_Busy;
Out_CYw_Rev_01_Pick_A_H := _p98;
Output_A_M[17] := _p98;
(* Rung 83 *)
_p99 := Output_A_M[17] AND TimerQ_In_SenCY_Rev_01_Pick_A_H;
Out_CYw_Rev_01_Pick_A_H_Done := _p99;
Output_A_Reset_TON[17](In := _p99, PT := T#1s);
(* Rung 84 *)
Output_A_Error_TON[17](In := Out_CYw_Rev_01_Pick_A_H_Auto[1] AND AutoMode AND NOT Pause[1] AND NOT TimerQ_In_SenCY_Rev_01_Pick_A_H, PT := T#10s);
_e100(CLK := Output_A_Error_TON[17].Q);
IF _e100.Q THEN
    Output_A_Error_M[17] := TRUE;
    HMI_MessageNo[0] := INT#23;
END_IF;

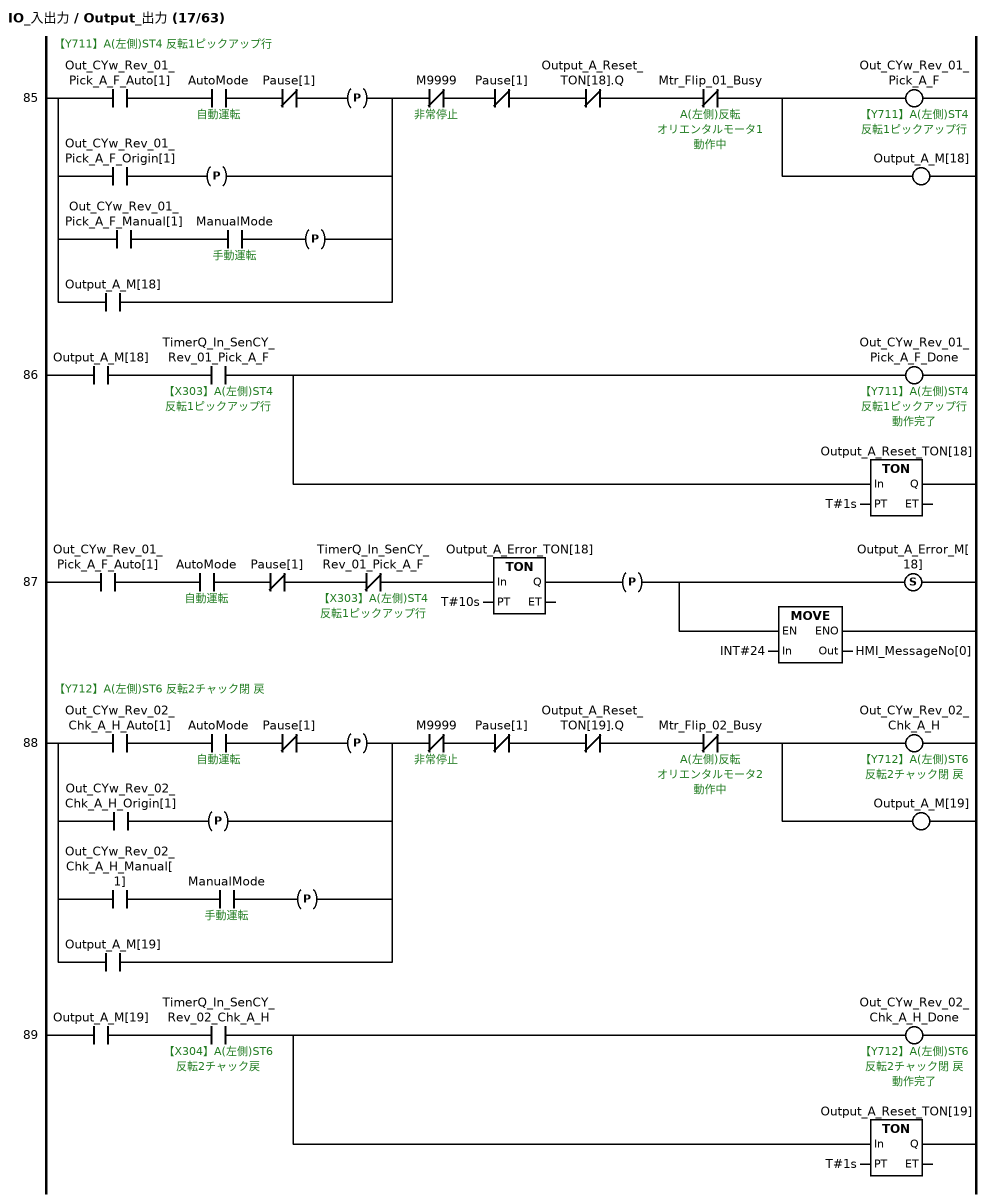
(* Rung 85: 【Y711】A(左側)ST4 反転1ピックアップ行 *)
_e101(CLK := Out_CYw_Rev_01_Pick_A_F_Auto[1] AND AutoMode AND NOT Pause[1]);
_e102(CLK := Out_CYw_Rev_01_Pick_A_F_Origin[1]);
_e103(CLK := Out_CYw_Rev_01_Pick_A_F_Manual[1] AND ManualMode);
_p104 := (_e101.Q OR _e102.Q OR _e103.Q OR Output_A_M[18]) AND NOT M9999 AND NOT Pause[1] AND NOT Output_A_Reset_TON[18].Q AND NOT Mtr_Flip_01_Busy;
Out_CYw_Rev_01_Pick_A_F := _p104;
Output_A_M[18] := _p104;
(* Rung 86 *)
_p105 := Output_A_M[18] AND TimerQ_In_SenCY_Rev_01_Pick_A_F;
Out_CYw_Rev_01_Pick_A_F_Done := _p105;
Output_A_Reset_TON[18](In := _p105, PT := T#1s);
(* Rung 87 *)
Output_A_Error_TON[18](In := Out_CYw_Rev_01_Pick_A_F_Auto[1] AND AutoMode AND NOT Pause[1] AND NOT TimerQ_In_SenCY_Rev_01_Pick_A_F, PT := T#10s);
_e106(CLK := Output_A_Error_TON[18].Q);
IF _e106.Q THEN
    Output_A_Error_M[18] := TRUE;
    HMI_MessageNo[0] := INT#24;
END_IF;
(* Rung 88: 【Y712】A(左側)ST6 反転2チャック閉 戻 *)
_e107(CLK := Out_CYw_Rev_02_Chk_A_H_Auto[1] AND AutoMode AND NOT Pause[1]);
_e108(CLK := Out_CYw_Rev_02_Chk_A_H_Origin[1]);
_e109(CLK := Out_CYw_Rev_02_Chk_A_H_Manual[1] AND ManualMode);
_p110 := (_e107.Q OR _e108.Q OR _e109.Q OR Output_A_M[19]) AND NOT M9999 AND NOT Pause[1] AND NOT Output_A_Reset_TON[19].Q AND NOT Mtr_Flip_02_Busy;
Out_CYw_Rev_02_Chk_A_H := _p110;
Output_A_M[19] := _p110;
(* Rung 89 *)
_p111 := Output_A_M[19] AND TimerQ_In_SenCY_Rev_02_Chk_A_H;
Out_CYw_Rev_02_Chk_A_H_Done := _p111;
Output_A_Reset_TON[19](In := _p111, PT := T#1s);

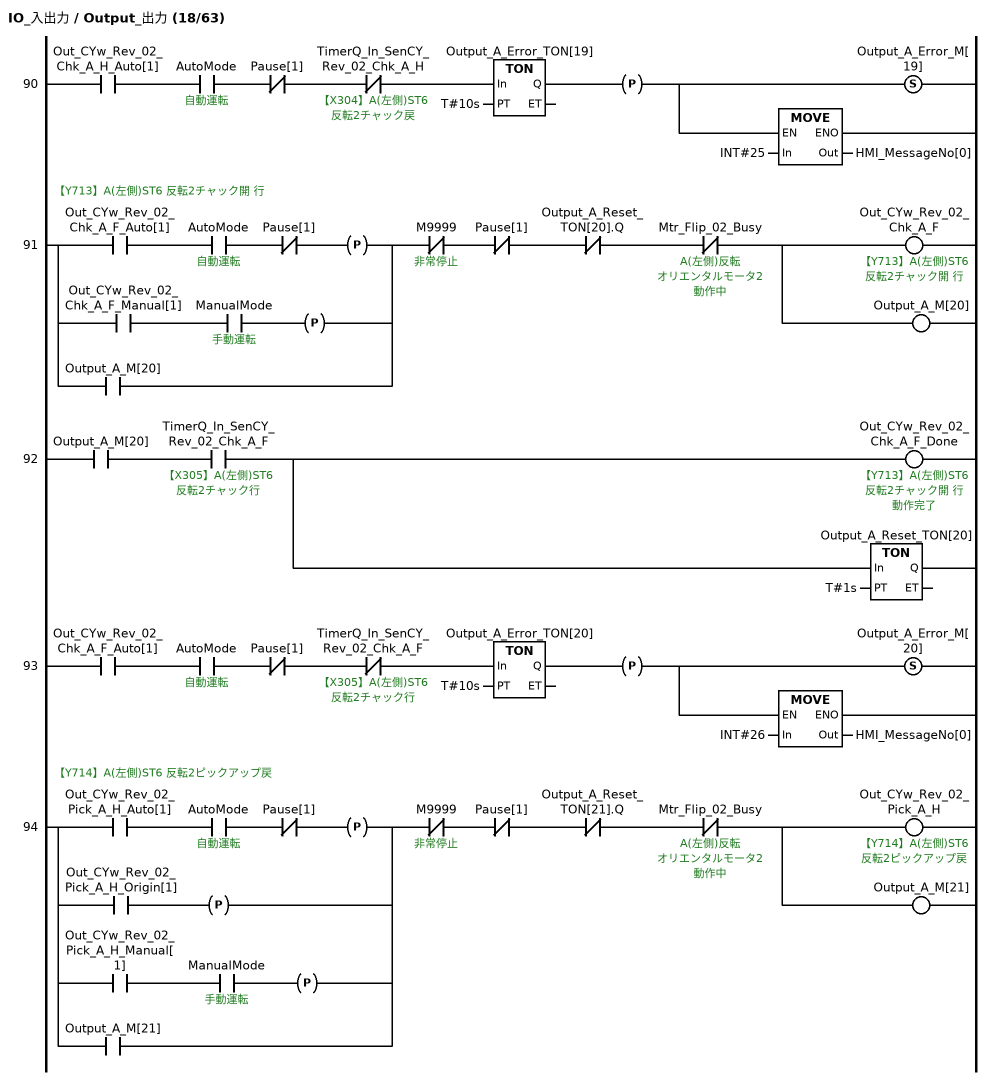
(* Rung 90 *)
Output_A_Error_TON[19](In := Out_CYw_Rev_02_Chk_A_H_Auto[1] AND AutoMode AND NOT Pause[1] AND NOT TimerQ_In_SenCY_Rev_02_Chk_A_H, PT := T#10s);
_e112(CLK := Output_A_Error_TON[19].Q);
IF _e112.Q THEN
    Output_A_Error_M[19] := TRUE;
    HMI_MessageNo[0] := INT#25;
END_IF;
(* Rung 91: 【Y713】A(左側)ST6 反転2チャック開 行 *)
_e113(CLK := Out_CYw_Rev_02_Chk_A_F_Auto[1] AND AutoMode AND NOT Pause[1]);
_e114(CLK := Out_CYw_Rev_02_Chk_A_F_Manual[1] AND ManualMode);
_p115 := (_e113.Q OR _e114.Q OR Output_A_M[20]) AND NOT M9999 AND NOT Pause[1] AND NOT Output_A_Reset_TON[20].Q AND NOT Mtr_Flip_02_Busy;
Out_CYw_Rev_02_Chk_A_F := _p115;
Output_A_M[20] := _p115;
(* Rung 92 *)
_p116 := Output_A_M[20] AND TimerQ_In_SenCY_Rev_02_Chk_A_F;
Out_CYw_Rev_02_Chk_A_F_Done := _p116;
Output_A_Reset_TON[20](In := _p116, PT := T#1s);
(* Rung 93 *)
Output_A_Error_TON[20](In := Out_CYw_Rev_02_Chk_A_F_Auto[1] AND AutoMode AND NOT Pause[1] AND NOT TimerQ_In_SenCY_Rev_02_Chk_A_F, PT := T#10s);
_e117(CLK := Output_A_Error_TON[20].Q);
IF _e117.Q THEN
    Output_A_Error_M[20] := TRUE;
    HMI_MessageNo[0] := INT#26;
END_IF;
(* Rung 94: 【Y714】A(左側)ST6 反転2ピックアップ戻 *)
_e118(CLK := Out_CYw_Rev_02_Pick_A_H_Auto[1] AND AutoMode AND NOT Pause[1]);
_e119(CLK := Out_CYw_Rev_02_Pick_A_H_Origin[1]);
_e120(CLK := Out_CYw_Rev_02_Pick_A_H_Manual[1] AND ManualMode);
_p121 := (_e118.Q OR _e119.Q OR _e120.Q OR Output_A_M[21]) AND NOT M9999 AND NOT Pause[1] AND NOT Output_A_Reset_TON[21].Q AND NOT Mtr_Flip_02_Busy;
Out_CYw_Rev_02_Pick_A_H := _p121;
Output_A_M[21] := _p121;

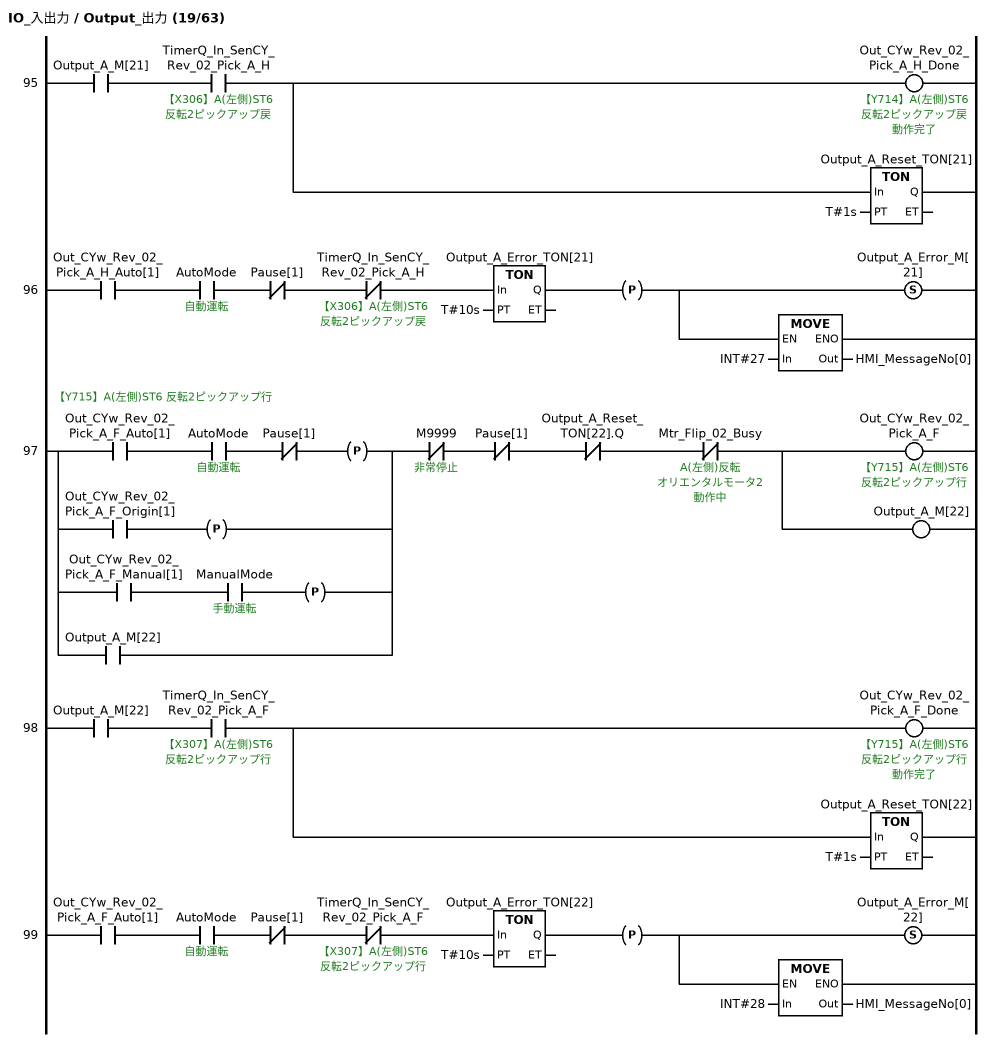
(* Rung 95 *)
_p122 := Output_A_M[21] AND TimerQ_In_SenCY_Rev_02_Pick_A_H;
Out_CYw_Rev_02_Pick_A_H_Done := _p122;
Output_A_Reset_TON[21](In := _p122, PT := T#1s);
(* Rung 96 *)
Output_A_Error_TON[21](In := Out_CYw_Rev_02_Pick_A_H_Auto[1] AND AutoMode AND NOT Pause[1] AND NOT TimerQ_In_SenCY_Rev_02_Pick_A_H, PT := T#10s);
_e123(CLK := Output_A_Error_TON[21].Q);
IF _e123.Q THEN
    Output_A_Error_M[21] := TRUE;
    HMI_MessageNo[0] := INT#27;
END_IF;
(* Rung 97: 【Y715】A(左側)ST6 反転2ピックアップ行 *)
_e124(CLK := Out_CYw_Rev_02_Pick_A_F_Auto[1] AND AutoMode AND NOT Pause[1]);
_e125(CLK := Out_CYw_Rev_02_Pick_A_F_Origin[1]);
_e126(CLK := Out_CYw_Rev_02_Pick_A_F_Manual[1] AND ManualMode);
_p127 := (_e124.Q OR _e125.Q OR _e126.Q OR Output_A_M[22]) AND NOT M9999 AND NOT Pause[1] AND NOT Output_A_Reset_TON[22].Q AND NOT Mtr_Flip_02_Busy;
Out_CYw_Rev_02_Pick_A_F := _p127;
Output_A_M[22] := _p127;
(* Rung 98 *)
_p128 := Output_A_M[22] AND TimerQ_In_SenCY_Rev_02_Pick_A_F;
Out_CYw_Rev_02_Pick_A_F_Done := _p128;
Output_A_Reset_TON[22](In := _p128, PT := T#1s);
(* Rung 99 *)
Output_A_Error_TON[22](In := Out_CYw_Rev_02_Pick_A_F_Auto[1] AND AutoMode AND NOT Pause[1] AND NOT TimerQ_In_SenCY_Rev_02_Pick_A_F, PT := T#10s);
_e129(CLK := Output_A_Error_TON[22].Q);
IF _e129.Q THEN
    Output_A_Error_M[22] := TRUE;
    HMI_MessageNo[0] := INT#28;
END_IF;

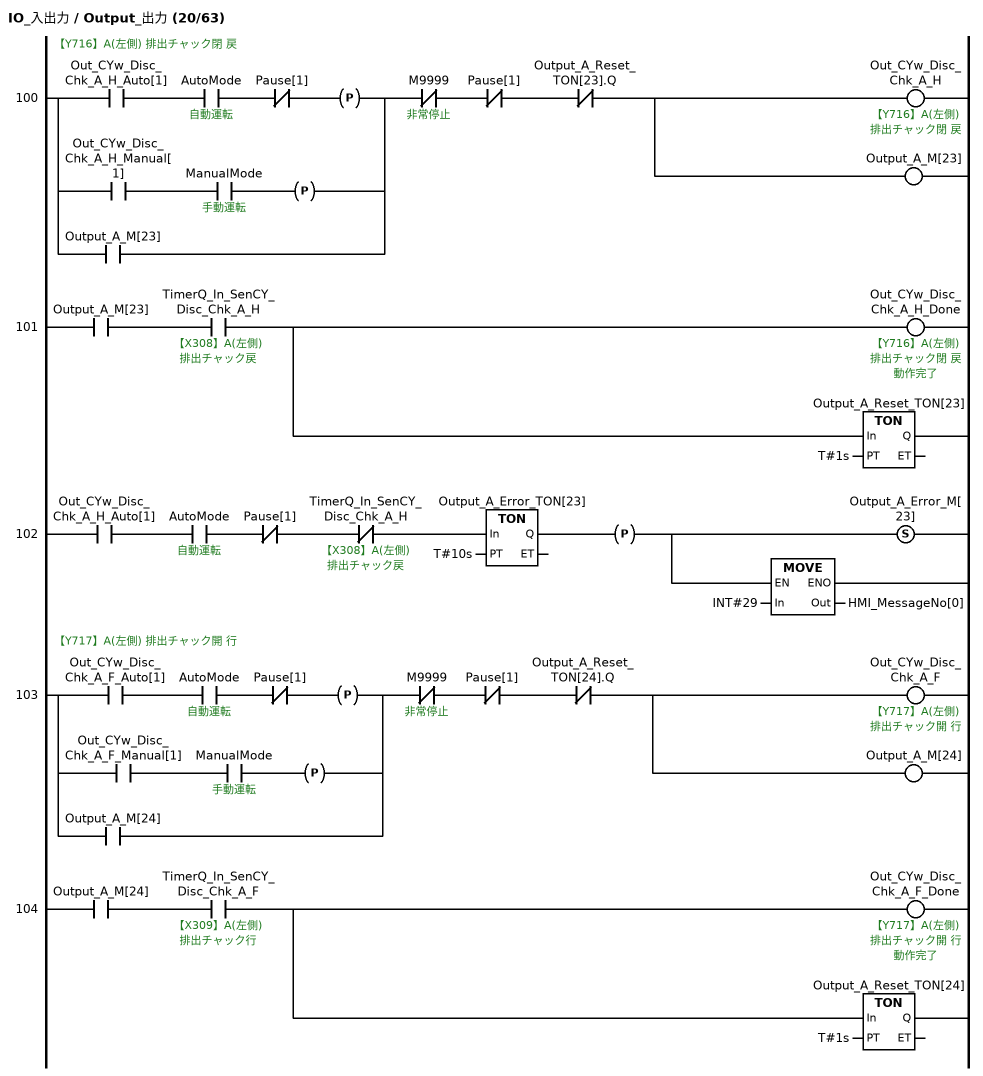
(* Rung 100: 【Y716】A(左側) 排出チャック閉 戻 *)
_e130(CLK := Out_CYw_Disc_Chk_A_H_Auto[1] AND AutoMode AND NOT Pause[1]);
_e131(CLK := Out_CYw_Disc_Chk_A_H_Manual[1] AND ManualMode);
_p132 := (_e130.Q OR _e131.Q OR Output_A_M[23]) AND NOT M9999 AND NOT Pause[1] AND NOT Output_A_Reset_TON[23].Q;
Out_CYw_Disc_Chk_A_H := _p132;
Output_A_M[23] := _p132;
(* Rung 101 *)
Out_CYw_Disc_Chk_A_H_Done := Output_A_M[23] AND TimerQ_In_SenCY_Disc_Chk_A_H;
Output_A_Reset_TON[23](In := Output_A_M[23] AND TimerQ_In_SenCY_Disc_Chk_A_H, PT := T#1s);
(* Rung 102 *)
Output_A_Error_TON[23](In := Out_CYw_Disc_Chk_A_H_Auto[1] AND AutoMode AND NOT Pause[1] AND NOT TimerQ_In_SenCY_Disc_Chk_A_H, PT := T#10s);
_e133(CLK := Output_A_Error_TON[23].Q);
IF _e133.Q THEN
    Output_A_Error_M[23] := TRUE;
    HMI_MessageNo[0] := INT#29;
END_IF;
(* Rung 103: 【Y717】A(左側) 排出チャック開 行 *)
_e134(CLK := Out_CYw_Disc_Chk_A_F_Auto[1] AND AutoMode AND NOT Pause[1]);
_e135(CLK := Out_CYw_Disc_Chk_A_F_Manual[1] AND ManualMode);
_p136 := (_e134.Q OR _e135.Q OR Output_A_M[24]) AND NOT M9999 AND NOT Pause[1] AND NOT Output_A_Reset_TON[24].Q;
Out_CYw_Disc_Chk_A_F := _p136;
Output_A_M[24] := _p136;
(* Rung 104 *)
Out_CYw_Disc_Chk_A_F_Done := Output_A_M[24] AND TimerQ_In_SenCY_Disc_Chk_A_F;
Output_A_Reset_TON[24](In := Output_A_M[24] AND TimerQ_In_SenCY_Disc_Chk_A_F, PT := T#1s);

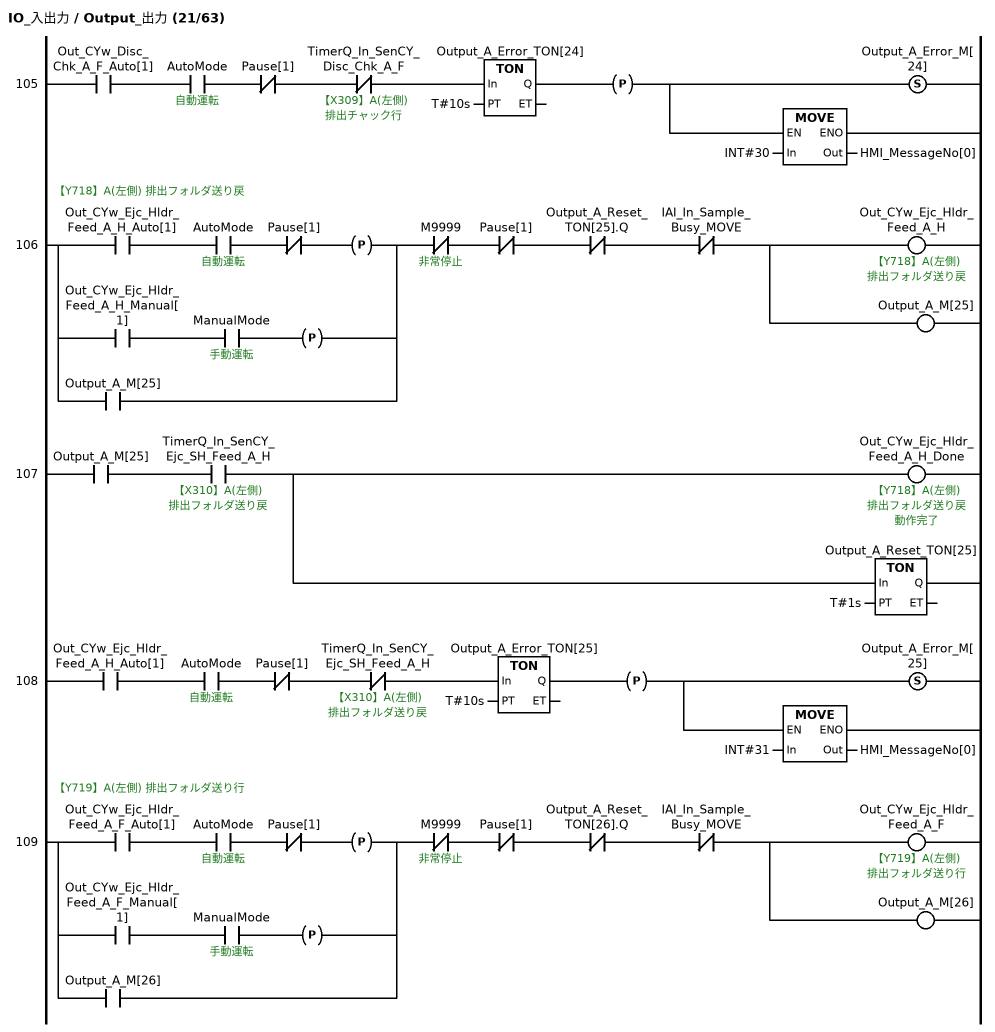
(* Rung 105 *)
Output_A_Error_TON[24](In := Out_CYw_Disc_Chk_A_F_Auto[1] AND AutoMode AND NOT Pause[1] AND NOT TimerQ_In_SenCY_Disc_Chk_A_F, PT := T#10s);
_e137(CLK := Output_A_Error_TON[24].Q);
IF _e137.Q THEN
    Output_A_Error_M[24] := TRUE;
    HMI_MessageNo[0] := INT#30;
END_IF;
(* Rung 106: 【Y718】A(左側) 排出フォルダ送り戻 *)
_e138(CLK := Out_CYw_Ejc_Hldr_Feed_A_H_Auto[1] AND AutoMode AND NOT Pause[1]);
_e139(CLK := Out_CYw_Ejc_Hldr_Feed_A_H_Manual[1] AND ManualMode);
_p140 := (_e138.Q OR _e139.Q OR Output_A_M[25]) AND NOT M9999 AND NOT Pause[1] AND NOT Output_A_Reset_TON[25].Q AND NOT IAI_In_Sample_Busy_MOVE;
Out_CYw_Ejc_Hldr_Feed_A_H := _p140;
Output_A_M[25] := _p140;
(* Rung 107 *)
_p141 := Output_A_M[25] AND TimerQ_In_SenCY_Ejc_SH_Feed_A_H;
Out_CYw_Ejc_Hldr_Feed_A_H_Done := _p141;
Output_A_Reset_TON[25](In := _p141, PT := T#1s);
(* Rung 108 *)
Output_A_Error_TON[25](In := Out_CYw_Ejc_Hldr_Feed_A_H_Auto[1] AND AutoMode AND NOT Pause[1] AND NOT TimerQ_In_SenCY_Ejc_SH_Feed_A_H, PT := T#10s);
_e142(CLK := Output_A_Error_TON[25].Q);
IF _e142.Q THEN
    Output_A_Error_M[25] := TRUE;
    HMI_MessageNo[0] := INT#31;
END_IF;
(* Rung 109: 【Y719】A(左側) 排出フォルダ送り行 *)
_e143(CLK := Out_CYw_Ejc_Hldr_Feed_A_F_Auto[1] AND AutoMode AND NOT Pause[1]);
_e144(CLK := Out_CYw_Ejc_Hldr_Feed_A_F_Manual[1] AND ManualMode);
_p145 := (_e143.Q OR _e144.Q OR Output_A_M[26]) AND NOT M9999 AND NOT Pause[1] AND NOT Output_A_Reset_TON[26].Q AND NOT IAI_In_Sample_Busy_MOVE;
Out_CYw_Ejc_Hldr_Feed_A_F := _p145;
Output_A_M[26] := _p145;

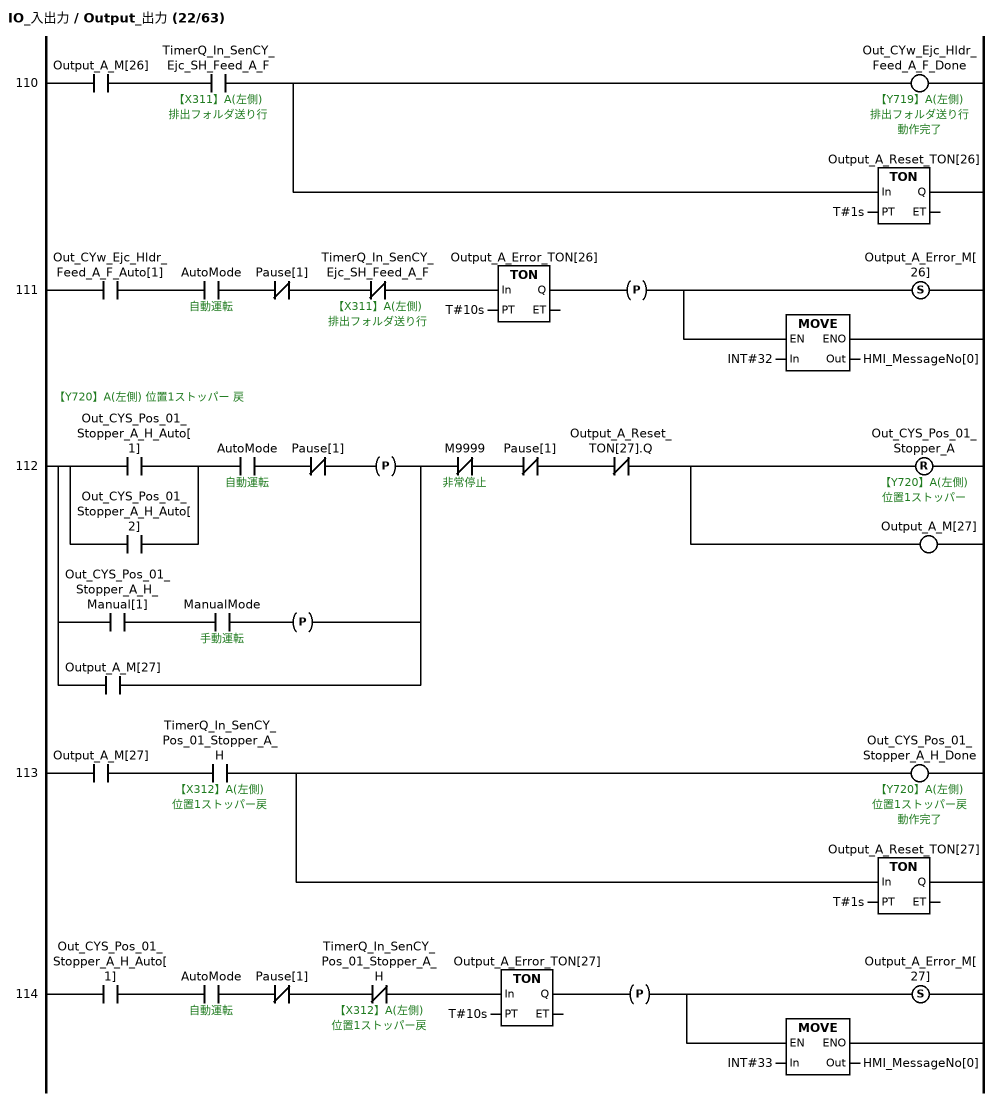
(* Rung 110 *)
_p146 := Output_A_M[26] AND TimerQ_In_SenCY_Ejc_SH_Feed_A_F;
Out_CYw_Ejc_Hldr_Feed_A_F_Done := _p146;
Output_A_Reset_TON[26](In := _p146, PT := T#1s);
(* Rung 111 *)
Output_A_Error_TON[26](In := Out_CYw_Ejc_Hldr_Feed_A_F_Auto[1] AND AutoMode AND NOT Pause[1] AND NOT TimerQ_In_SenCY_Ejc_SH_Feed_A_F, PT := T#10s);
_e147(CLK := Output_A_Error_TON[26].Q);
IF _e147.Q THEN
    Output_A_Error_M[26] := TRUE;
    HMI_MessageNo[0] := INT#32;
END_IF;
(* Rung 112: 【Y720】A(左側) 位置1ストッパー 戻 *)
_e148(CLK := (Out_CYS_Pos_01_Stopper_A_H_Auto[1] OR Out_CYS_Pos_01_Stopper_A_H_Auto[2]) AND AutoMode AND NOT Pause[1]);
_e149(CLK := Out_CYS_Pos_01_Stopper_A_H_Manual[1] AND ManualMode);
_p150 := (_e148.Q OR _e149.Q OR Output_A_M[27]) AND NOT M9999 AND NOT Pause[1] AND NOT Output_A_Reset_TON[27].Q;
IF _p150 THEN Out_CYS_Pos_01_Stopper_A := FALSE; END_IF;
Output_A_M[27] := _p150;
(* Rung 113 *)
_p151 := Output_A_M[27] AND TimerQ_In_SenCY_Pos_01_Stopper_A_H;
Out_CYS_Pos_01_Stopper_A_H_Done := _p151;
Output_A_Reset_TON[27](In := _p151, PT := T#1s);
(* Rung 114 *)
Output_A_Error_TON[27](In := Out_CYS_Pos_01_Stopper_A_H_Auto[1] AND AutoMode AND NOT Pause[1] AND NOT TimerQ_In_SenCY_Pos_01_Stopper_A_H, PT := T#10s);
_e152(CLK := Output_A_Error_TON[27].Q);
IF _e152.Q THEN
    Output_A_Error_M[27] := TRUE;
    HMI_MessageNo[0] := INT#33;
END_IF;

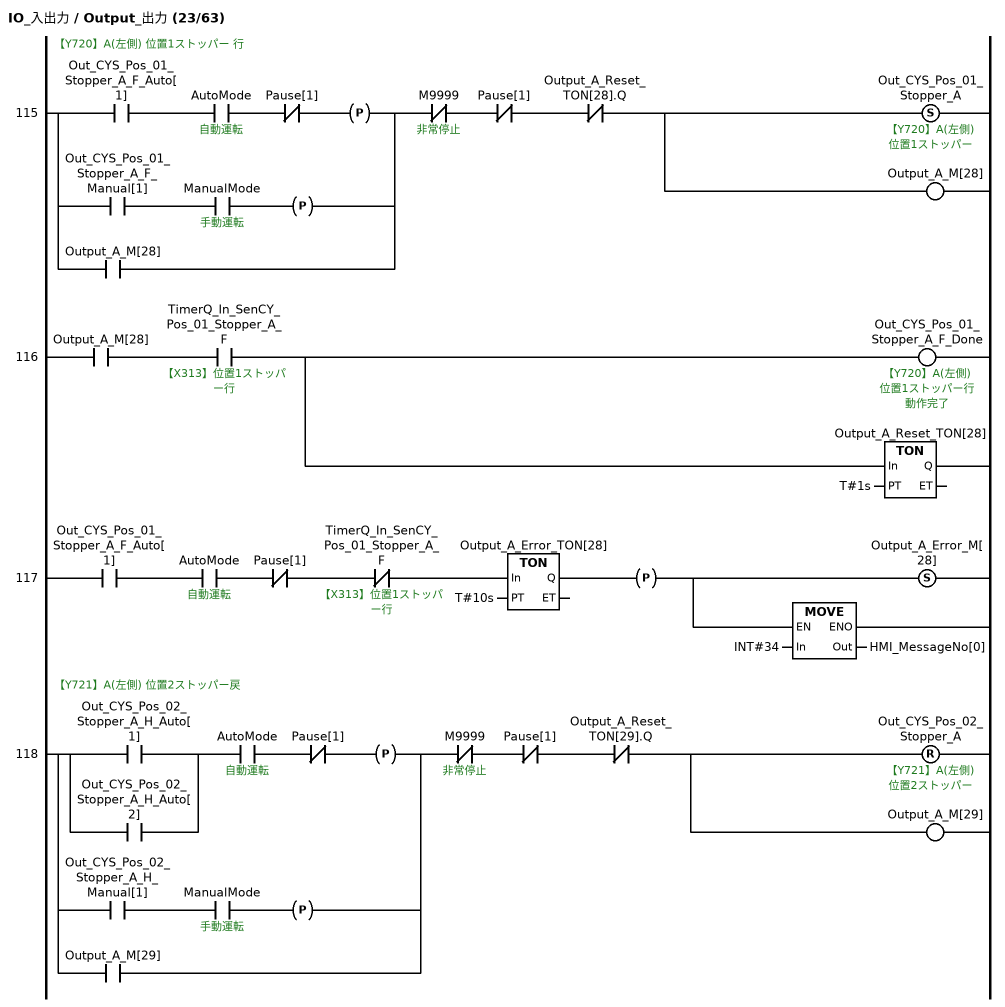
(* Rung 115: 【Y720】A(左側) 位置1ストッパー 行 *)
_e153(CLK := Out_CYS_Pos_01_Stopper_A_F_Auto[1] AND AutoMode AND NOT Pause[1]);
_e154(CLK := Out_CYS_Pos_01_Stopper_A_F_Manual[1] AND ManualMode);
_p155 := (_e153.Q OR _e154.Q OR Output_A_M[28]) AND NOT M9999 AND NOT Pause[1] AND NOT Output_A_Reset_TON[28].Q;
IF _p155 THEN Out_CYS_Pos_01_Stopper_A := TRUE; END_IF;
Output_A_M[28] := _p155;
(* Rung 116 *)
_p156 := Output_A_M[28] AND TimerQ_In_SenCY_Pos_01_Stopper_A_F;
Out_CYS_Pos_01_Stopper_A_F_Done := _p156;
Output_A_Reset_TON[28](In := _p156, PT := T#1s);
(* Rung 117 *)
Output_A_Error_TON[28](In := Out_CYS_Pos_01_Stopper_A_F_Auto[1] AND AutoMode AND NOT Pause[1] AND NOT TimerQ_In_SenCY_Pos_01_Stopper_A_F, PT := T#10s);
_e157(CLK := Output_A_Error_TON[28].Q);
IF _e157.Q THEN
    Output_A_Error_M[28] := TRUE;
    HMI_MessageNo[0] := INT#34;
END_IF;
(* Rung 118: 【Y721】A(左側) 位置2ストッパー戻 *)
_e158(CLK := (Out_CYS_Pos_02_Stopper_A_H_Auto[1] OR Out_CYS_Pos_02_Stopper_A_H_Auto[2]) AND AutoMode AND NOT Pause[1]);
_e159(CLK := Out_CYS_Pos_02_Stopper_A_H_Manual[1] AND ManualMode);
_p160 := (_e158.Q OR _e159.Q OR Output_A_M[29]) AND NOT M9999 AND NOT Pause[1] AND NOT Output_A_Reset_TON[29].Q;
IF _p160 THEN Out_CYS_Pos_02_Stopper_A := FALSE; END_IF;
Output_A_M[29] := _p160;

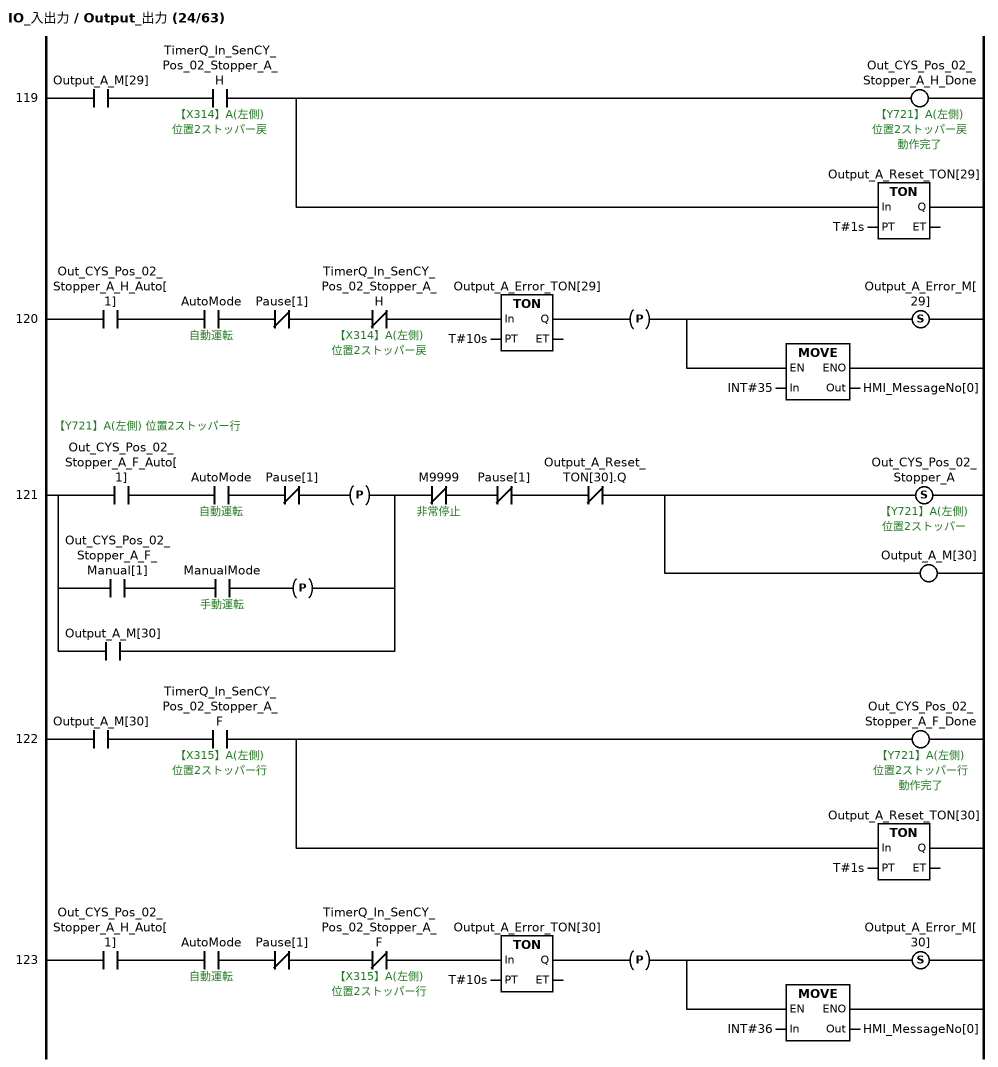
(* Rung 119 *)
_p161 := Output_A_M[29] AND TimerQ_In_SenCY_Pos_02_Stopper_A_H;
Out_CYS_Pos_02_Stopper_A_H_Done := _p161;
Output_A_Reset_TON[29](In := _p161, PT := T#1s);
(* Rung 120 *)
Output_A_Error_TON[29](In := Out_CYS_Pos_02_Stopper_A_H_Auto[1] AND AutoMode AND NOT Pause[1] AND NOT TimerQ_In_SenCY_Pos_02_Stopper_A_H, PT := T#10s);
_e162(CLK := Output_A_Error_TON[29].Q);
IF _e162.Q THEN
    Output_A_Error_M[29] := TRUE;
    HMI_MessageNo[0] := INT#35;
END_IF;
(* Rung 121: 【Y721】A(左側) 位置2ストッパー行 *)
_e163(CLK := Out_CYS_Pos_02_Stopper_A_F_Auto[1] AND AutoMode AND NOT Pause[1]);
_e164(CLK := Out_CYS_Pos_02_Stopper_A_F_Manual[1] AND ManualMode);
_p165 := (_e163.Q OR _e164.Q OR Output_A_M[30]) AND NOT M9999 AND NOT Pause[1] AND NOT Output_A_Reset_TON[30].Q;
IF _p165 THEN Out_CYS_Pos_02_Stopper_A := TRUE; END_IF;
Output_A_M[30] := _p165;
(* Rung 122 *)
_p166 := Output_A_M[30] AND TimerQ_In_SenCY_Pos_02_Stopper_A_F;
Out_CYS_Pos_02_Stopper_A_F_Done := _p166;
Output_A_Reset_TON[30](In := _p166, PT := T#1s);
(* Rung 123 *)
Output_A_Error_TON[30](In := Out_CYS_Pos_02_Stopper_A_H_Auto[1] AND AutoMode AND NOT Pause[1] AND NOT TimerQ_In_SenCY_Pos_02_Stopper_A_F, PT := T#10s);
_e167(CLK := Output_A_Error_TON[30].Q);
IF _e167.Q THEN
    Output_A_Error_M[30] := TRUE;
    HMI_MessageNo[0] := INT#36;
END_IF;

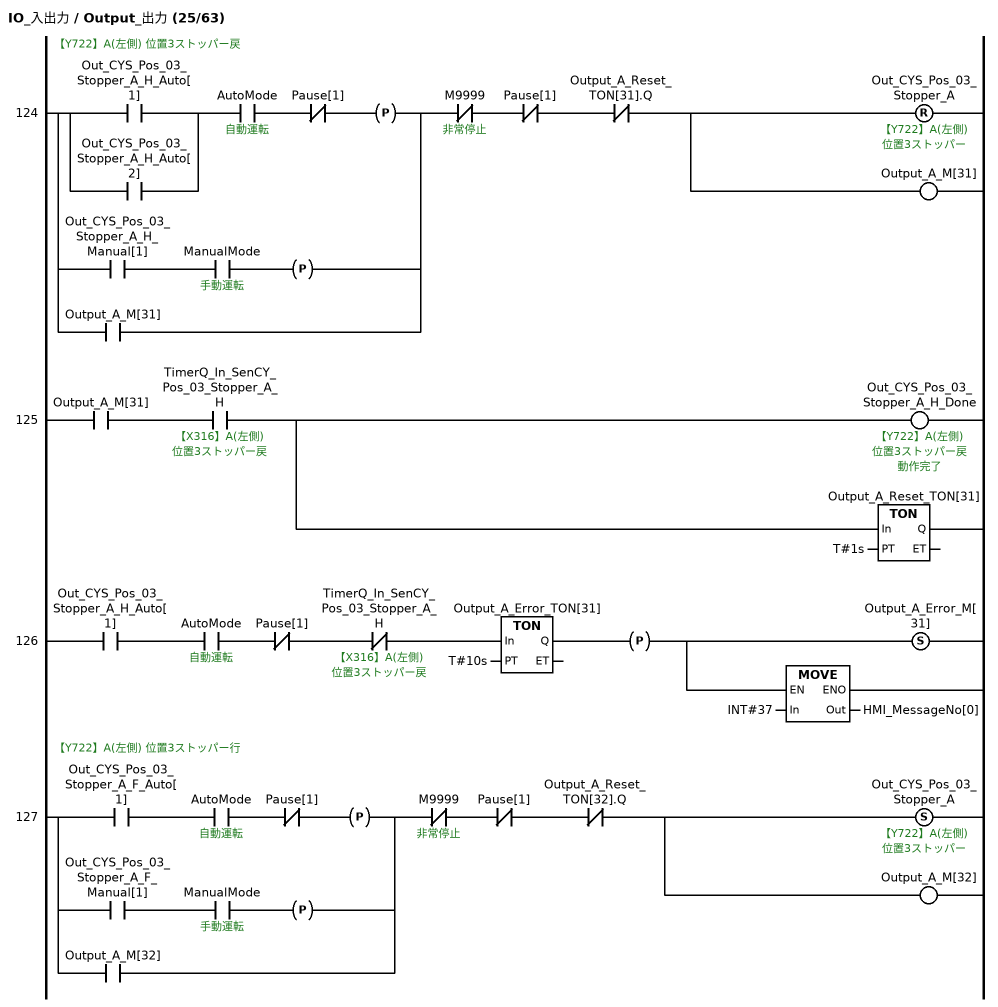
(* Rung 124: 【Y722】A(左側) 位置3ストッパー戻 *)
_e168(CLK := (Out_CYS_Pos_03_Stopper_A_H_Auto[1] OR Out_CYS_Pos_03_Stopper_A_H_Auto[2]) AND AutoMode AND NOT Pause[1]);
_e169(CLK := Out_CYS_Pos_03_Stopper_A_H_Manual[1] AND ManualMode);
_p170 := (_e168.Q OR _e169.Q OR Output_A_M[31]) AND NOT M9999 AND NOT Pause[1] AND NOT Output_A_Reset_TON[31].Q;
IF _p170 THEN Out_CYS_Pos_03_Stopper_A := FALSE; END_IF;
Output_A_M[31] := _p170;
(* Rung 125 *)
_p171 := Output_A_M[31] AND TimerQ_In_SenCY_Pos_03_Stopper_A_H;
Out_CYS_Pos_03_Stopper_A_H_Done := _p171;
Output_A_Reset_TON[31](In := _p171, PT := T#1s);
(* Rung 126 *)
Output_A_Error_TON[31](In := Out_CYS_Pos_03_Stopper_A_H_Auto[1] AND AutoMode AND NOT Pause[1] AND NOT TimerQ_In_SenCY_Pos_03_Stopper_A_H, PT := T#10s);
_e172(CLK := Output_A_Error_TON[31].Q);
IF _e172.Q THEN
    Output_A_Error_M[31] := TRUE;
    HMI_MessageNo[0] := INT#37;
END_IF;
(* Rung 127: 【Y722】A(左側) 位置3ストッパー行 *)
_e173(CLK := Out_CYS_Pos_03_Stopper_A_F_Auto[1] AND AutoMode AND NOT Pause[1]);
_e174(CLK := Out_CYS_Pos_03_Stopper_A_F_Manual[1] AND ManualMode);
_p175 := (_e173.Q OR _e174.Q OR Output_A_M[32]) AND NOT M9999 AND NOT Pause[1] AND NOT Output_A_Reset_TON[32].Q;
IF _p175 THEN Out_CYS_Pos_03_Stopper_A := TRUE; END_IF;
Output_A_M[32] := _p175;

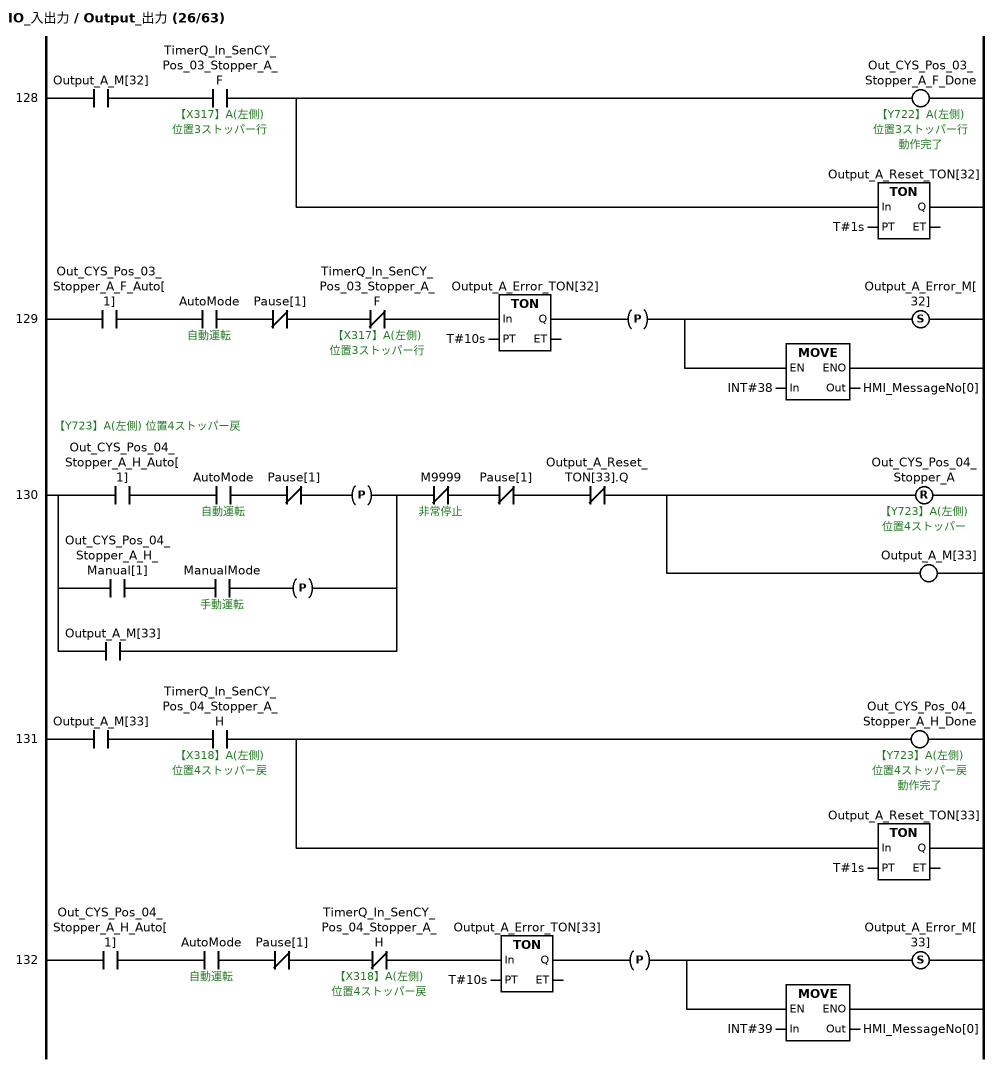
(* Rung 128 *)
_p176 := Output_A_M[32] AND TimerQ_In_SenCY_Pos_03_Stopper_A_F;
Out_CYS_Pos_03_Stopper_A_F_Done := _p176;
Output_A_Reset_TON[32](In := _p176, PT := T#1s);
(* Rung 129 *)
Output_A_Error_TON[32](In := Out_CYS_Pos_03_Stopper_A_F_Auto[1] AND AutoMode AND NOT Pause[1] AND NOT TimerQ_In_SenCY_Pos_03_Stopper_A_F, PT := T#10s);
_e177(CLK := Output_A_Error_TON[32].Q);
IF _e177.Q THEN
    Output_A_Error_M[32] := TRUE;
    HMI_MessageNo[0] := INT#38;
END_IF;
(* Rung 130: 【Y723】A(左側) 位置4ストッパー戻 *)
_e178(CLK := Out_CYS_Pos_04_Stopper_A_H_Auto[1] AND AutoMode AND NOT Pause[1]);
_e179(CLK := Out_CYS_Pos_04_Stopper_A_H_Manual[1] AND ManualMode);
_p180 := (_e178.Q OR _e179.Q OR Output_A_M[33]) AND NOT M9999 AND NOT Pause[1] AND NOT Output_A_Reset_TON[33].Q;
IF _p180 THEN Out_CYS_Pos_04_Stopper_A := FALSE; END_IF;
Output_A_M[33] := _p180;
(* Rung 131 *)
_p181 := Output_A_M[33] AND TimerQ_In_SenCY_Pos_04_Stopper_A_H;
Out_CYS_Pos_04_Stopper_A_H_Done := _p181;
Output_A_Reset_TON[33](In := _p181, PT := T#1s);
(* Rung 132 *)
Output_A_Error_TON[33](In := Out_CYS_Pos_04_Stopper_A_H_Auto[1] AND AutoMode AND NOT Pause[1] AND NOT TimerQ_In_SenCY_Pos_04_Stopper_A_H, PT := T#10s);
_e182(CLK := Output_A_Error_TON[33].Q);
IF _e182.Q THEN
    Output_A_Error_M[33] := TRUE;
    HMI_MessageNo[0] := INT#39;
END_IF;

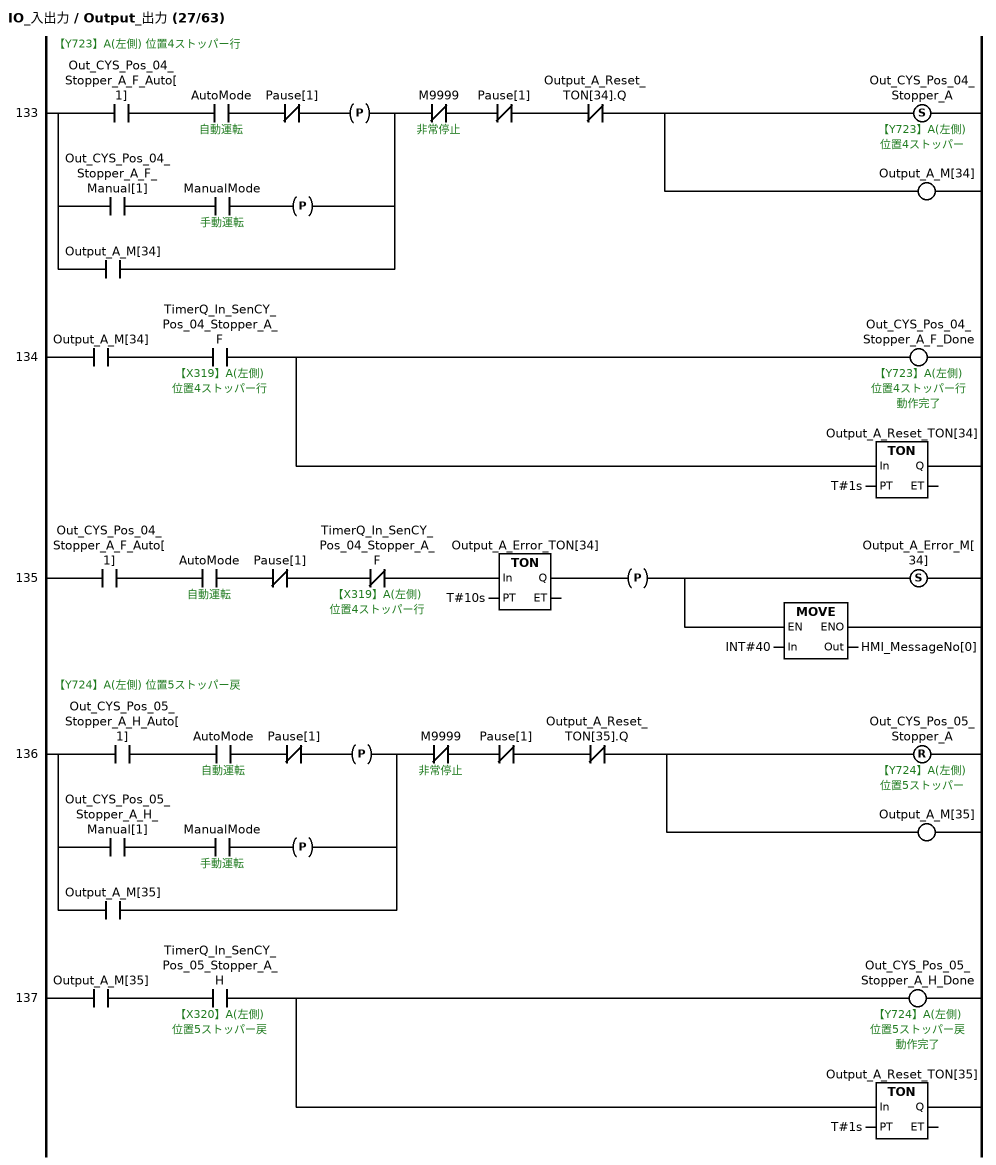
(* Rung 133: 【Y723】A(左側) 位置4ストッパー行 *)
_e183(CLK := Out_CYS_Pos_04_Stopper_A_F_Auto[1] AND AutoMode AND NOT Pause[1]);
_e184(CLK := Out_CYS_Pos_04_Stopper_A_F_Manual[1] AND ManualMode);
_p185 := (_e183.Q OR _e184.Q OR Output_A_M[34]) AND NOT M9999 AND NOT Pause[1] AND NOT Output_A_Reset_TON[34].Q;
IF _p185 THEN Out_CYS_Pos_04_Stopper_A := TRUE; END_IF;
Output_A_M[34] := _p185;
(* Rung 134 *)
_p186 := Output_A_M[34] AND TimerQ_In_SenCY_Pos_04_Stopper_A_F;
Out_CYS_Pos_04_Stopper_A_F_Done := _p186;
Output_A_Reset_TON[34](In := _p186, PT := T#1s);
(* Rung 135 *)
Output_A_Error_TON[34](In := Out_CYS_Pos_04_Stopper_A_F_Auto[1] AND AutoMode AND NOT Pause[1] AND NOT TimerQ_In_SenCY_Pos_04_Stopper_A_F, PT := T#10s);
_e187(CLK := Output_A_Error_TON[34].Q);
IF _e187.Q THEN
    Output_A_Error_M[34] := TRUE;
    HMI_MessageNo[0] := INT#40;
END_IF;
(* Rung 136: 【Y724】A(左側) 位置5ストッパー戻 *)
_e188(CLK := Out_CYS_Pos_05_Stopper_A_H_Auto[1] AND AutoMode AND NOT Pause[1]);
_e189(CLK := Out_CYS_Pos_05_Stopper_A_H_Manual[1] AND ManualMode);
_p190 := (_e188.Q OR _e189.Q OR Output_A_M[35]) AND NOT M9999 AND NOT Pause[1] AND NOT Output_A_Reset_TON[35].Q;
IF _p190 THEN Out_CYS_Pos_05_Stopper_A := FALSE; END_IF;
Output_A_M[35] := _p190;
(* Rung 137 *)
_p191 := Output_A_M[35] AND TimerQ_In_SenCY_Pos_05_Stopper_A_H;
Out_CYS_Pos_05_Stopper_A_H_Done := _p191;
Output_A_Reset_TON[35](In := _p191, PT := T#1s);

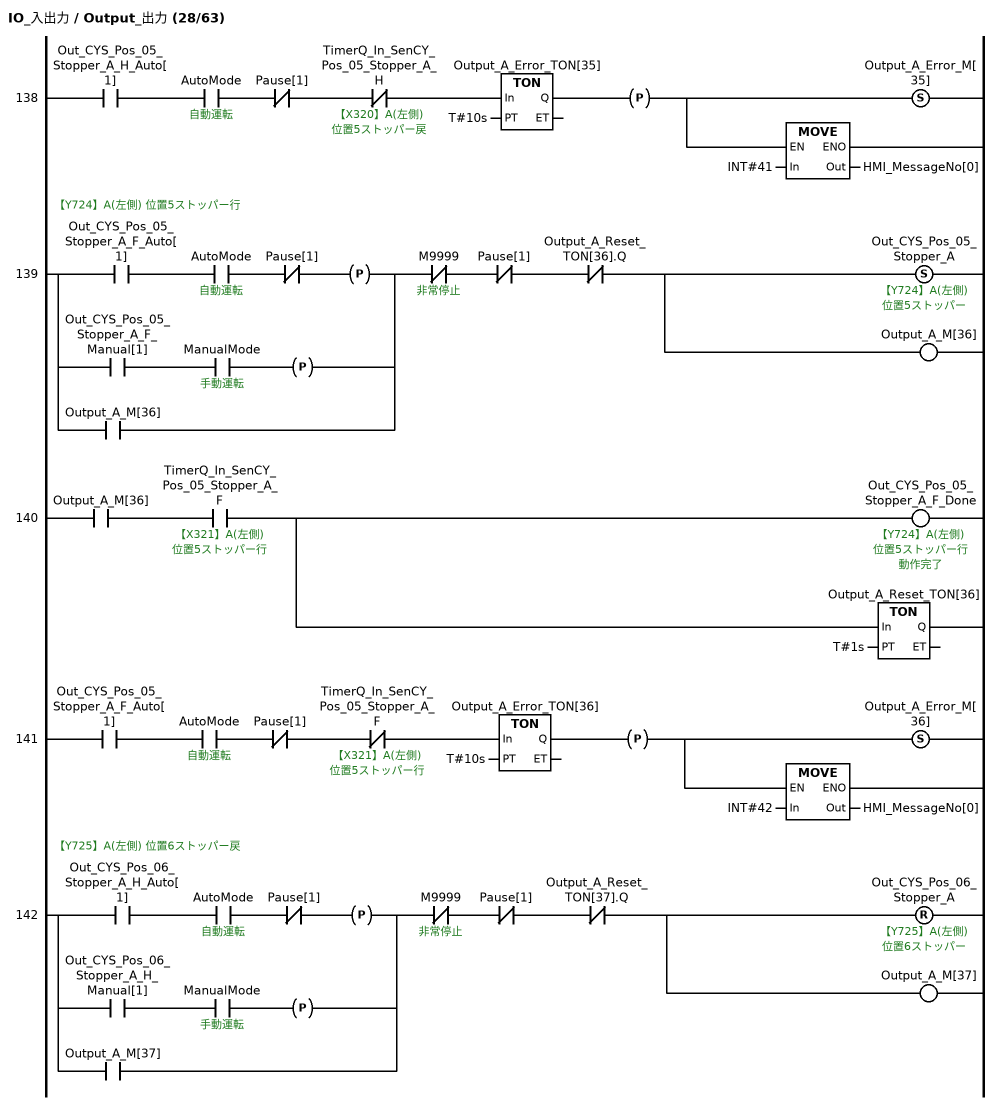
(* Rung 138 *)
Output_A_Error_TON[35](In := Out_CYS_Pos_05_Stopper_A_H_Auto[1] AND AutoMode AND NOT Pause[1] AND NOT TimerQ_In_SenCY_Pos_05_Stopper_A_H, PT := T#10s);
_e192(CLK := Output_A_Error_TON[35].Q);
IF _e192.Q THEN
    Output_A_Error_M[35] := TRUE;
    HMI_MessageNo[0] := INT#41;
END_IF;
(* Rung 139: 【Y724】A(左側) 位置5ストッパー行 *)
_e193(CLK := Out_CYS_Pos_05_Stopper_A_F_Auto[1] AND AutoMode AND NOT Pause[1]);
_e194(CLK := Out_CYS_Pos_05_Stopper_A_F_Manual[1] AND ManualMode);
_p195 := (_e193.Q OR _e194.Q OR Output_A_M[36]) AND NOT M9999 AND NOT Pause[1] AND NOT Output_A_Reset_TON[36].Q;
IF _p195 THEN Out_CYS_Pos_05_Stopper_A := TRUE; END_IF;
Output_A_M[36] := _p195;
(* Rung 140 *)
_p196 := Output_A_M[36] AND TimerQ_In_SenCY_Pos_05_Stopper_A_F;
Out_CYS_Pos_05_Stopper_A_F_Done := _p196;
Output_A_Reset_TON[36](In := _p196, PT := T#1s);
(* Rung 141 *)
Output_A_Error_TON[36](In := Out_CYS_Pos_05_Stopper_A_F_Auto[1] AND AutoMode AND NOT Pause[1] AND NOT TimerQ_In_SenCY_Pos_05_Stopper_A_F, PT := T#10s);
_e197(CLK := Output_A_Error_TON[36].Q);
IF _e197.Q THEN
    Output_A_Error_M[36] := TRUE;
    HMI_MessageNo[0] := INT#42;
END_IF;
(* Rung 142: 【Y725】A(左側) 位置6ストッパー戻 *)
_e198(CLK := Out_CYS_Pos_06_Stopper_A_H_Auto[1] AND AutoMode AND NOT Pause[1]);
_e199(CLK := Out_CYS_Pos_06_Stopper_A_H_Manual[1] AND ManualMode);
_p200 := (_e198.Q OR _e199.Q OR Output_A_M[37]) AND NOT M9999 AND NOT Pause[1] AND NOT Output_A_Reset_TON[37].Q;
IF _p200 THEN Out_CYS_Pos_06_Stopper_A := FALSE; END_IF;
Output_A_M[37] := _p200;

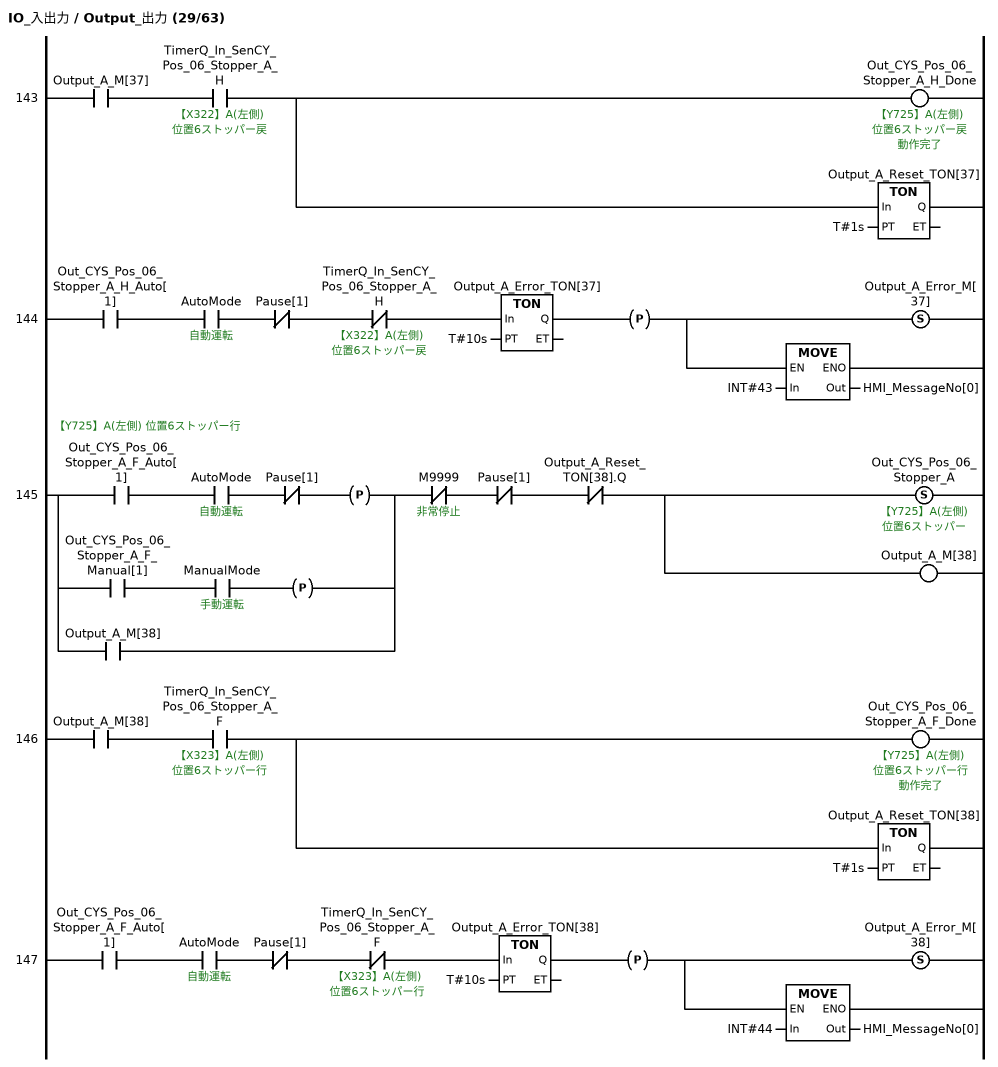
(* Rung 143 *)
_p201 := Output_A_M[37] AND TimerQ_In_SenCY_Pos_06_Stopper_A_H;
Out_CYS_Pos_06_Stopper_A_H_Done := _p201;
Output_A_Reset_TON[37](In := _p201, PT := T#1s);
(* Rung 144 *)
Output_A_Error_TON[37](In := Out_CYS_Pos_06_Stopper_A_H_Auto[1] AND AutoMode AND NOT Pause[1] AND NOT TimerQ_In_SenCY_Pos_06_Stopper_A_H, PT := T#10s);
_e202(CLK := Output_A_Error_TON[37].Q);
IF _e202.Q THEN
    Output_A_Error_M[37] := TRUE;
    HMI_MessageNo[0] := INT#43;
END_IF;
(* Rung 145: 【Y725】A(左側) 位置6ストッパー行 *)
_e203(CLK := Out_CYS_Pos_06_Stopper_A_F_Auto[1] AND AutoMode AND NOT Pause[1]);
_e204(CLK := Out_CYS_Pos_06_Stopper_A_F_Manual[1] AND ManualMode);
_p205 := (_e203.Q OR _e204.Q OR Output_A_M[38]) AND NOT M9999 AND NOT Pause[1] AND NOT Output_A_Reset_TON[38].Q;
IF _p205 THEN Out_CYS_Pos_06_Stopper_A := TRUE; END_IF;
Output_A_M[38] := _p205;
(* Rung 146 *)
_p206 := Output_A_M[38] AND TimerQ_In_SenCY_Pos_06_Stopper_A_F;
Out_CYS_Pos_06_Stopper_A_F_Done := _p206;
Output_A_Reset_TON[38](In := _p206, PT := T#1s);
(* Rung 147 *)
Output_A_Error_TON[38](In := Out_CYS_Pos_06_Stopper_A_F_Auto[1] AND AutoMode AND NOT Pause[1] AND NOT TimerQ_In_SenCY_Pos_06_Stopper_A_F, PT := T#10s);
_e207(CLK := Output_A_Error_TON[38].Q);
IF _e207.Q THEN
    Output_A_Error_M[38] := TRUE;
    HMI_MessageNo[0] := INT#44;
END_IF;

